{attribute 'external_name' := 'cmp_rts_DFC_rbr_safoutChnl3'}
TYPE DFC_rbr_safoutChnl3 : STRUCT
  DTC : UDINT := 16#200A00;
  DFCid : UINT := 802;
  debounceMethod : USINT := NO_DEBOUNCE;
END_STRUCT;
END_TYPE

{attribute 'external_name' := 'cmp_rts_DFC_rbr_safoutChnl4'}
TYPE DFC_rbr_safoutChnl4 : STRUCT
  DTC : UDINT := 16#200B00;
  DFCid : UINT := 805;
  debounceMethod : USINT := NO_DEBOUNCE;
END_STRUCT;
END_TYPE

{attribute 'external_name' := 'cmp_rts_DFC_rbr_safoutChnl5'}
TYPE DFC_rbr_safoutChnl5 : STRUCT
  DTC : UDINT := 16#200C00;
  DFCid : UINT := 808;
  debounceMethod : USINT := NO_DEBOUNCE;
END_STRUCT;
END_TYPE

{attribute 'external_name' := 'cmp_rts_DFC_rbr_safoutChnl6'}
TYPE DFC_rbr_safoutChnl6 : STRUCT
  DTC : UDINT := 16#201900;
  DFCid : UINT := 811;
  debounceMethod : USINT := NO_DEBOUNCE;
END_STRUCT;
END_TYPE

{attribute 'external_name' := 'cmp_rts_DFC_rbr_safoutChnl7'}
TYPE DFC_rbr_safoutChnl7 : STRUCT
  DTC : UDINT := 16#201A00;
  DFCid : UINT := 814;
  debounceMethod : USINT := NO_DEBOUNCE;
END_STRUCT;
END_TYPE

{attribute 'external_name' := 'cmp_rts_DFC_rbr_safoutChnl8'}
TYPE DFC_rbr_safoutChnl8 : STRUCT
  DTC : UDINT := 16#201B00;
  DFCid : UINT := 817;
  debounceMethod : USINT := NO_DEBOUNCE;
END_STRUCT;
END_TYPE

{attribute 'external_name' := 'cmp_rts_DFC_rbr_safoutChnl9'}
TYPE DFC_rbr_safoutChnl9 : STRUCT
  DTC : UDINT := 16#201C00;
  DFCid : UINT := 820;
  debounceMethod : USINT := NO_DEBOUNCE;
END_STRUCT;
END_TYPE

{attribute 'external_name' := 'cmp_rts_DFC_rbr_safoutChnl10'}
TYPE DFC_rbr_safoutChnl10 : STRUCT
  DTC : UDINT := 16#201D00;
  DFCid : UINT := 770;
  debounceMethod : USINT := NO_DEBOUNCE;
END_STRUCT;
END_TYPE

{attribute 'external_name' := 'cmp_rts_DFC_rbr_safoutChnl11'}
TYPE DFC_rbr_safoutChnl11 : STRUCT
  DTC : UDINT := 16#201E00;
  DFCid : UINT := 773;
  debounceMethod : USINT := NO_DEBOUNCE;
END_STRUCT;
END_TYPE

{attribute 'external_name' := 'cmp_rts_DFC_rbr_safoutChnl12'}
TYPE DFC_rbr_safoutChnl12 : STRUCT
  DTC : UDINT := 16#201F00;
  DFCid : UINT := 776;
  debounceMethod : USINT := NO_DEBOUNCE;
END_STRUCT;
END_TYPE

{attribute 'external_name' := 'cmp_rts_DFC_rbr_safoutChnl13'}
TYPE DFC_rbr_safoutChnl13 : STRUCT
  DTC : UDINT := 16#202000;
  DFCid : UINT := 779;
  debounceMethod : USINT := NO_DEBOUNCE;
END_STRUCT;
END_TYPE

{attribute 'external_name' := 'cmp_rts_DFC_rbr_safoutChnl14'}
TYPE DFC_rbr_safoutChnl14 : STRUCT
  DTC : UDINT := 16#202100;
  DFCid : UINT := 782;
  debounceMethod : USINT := NO_DEBOUNCE;
END_STRUCT;
END_TYPE

{attribute 'external_name' := 'cmp_rts_DFC_rbr_safoutChnl15'}
TYPE DFC_rbr_safoutChnl15 : STRUCT
  DTC : UDINT := 16#202200;
  DFCid : UINT := 785;
  debounceMethod : USINT := NO_DEBOUNCE;
END_STRUCT;
END_TYPE

{attribute 'external_name' := 'cmp_rts_DFC_rbr_safoutChnl16'}
TYPE DFC_rbr_safoutChnl16 : STRUCT
  DTC : UDINT := 16#202300;
  DFCid : UINT := 788;
  debounceMethod : USINT := NO_DEBOUNCE;
END_STRUCT;
END_TYPE

{attribute 'external_name' := 'cmp_rts_DFC_rbr_safoutChnl17'}
TYPE DFC_rbr_safoutChnl17 : STRUCT
  DTC : UDINT := 16#202400;
  DFCid : UINT := 791;
  debounceMethod : USINT := NO_DEBOUNCE;
END_STRUCT;
END_TYPE

{attribute 'external_name' := 'cmp_rts_DFC_rbr_safoutChnl18'}
TYPE DFC_rbr_safoutChnl18 : STRUCT
  DTC : UDINT := 16#202500;
  DFCid : UINT := 794;
  debounceMethod : USINT := NO_DEBOUNCE;
END_STRUCT;
END_TYPE

{attribute 'external_name' := 'cmp_rts_DFC_rbr_safoutChnl6Dev'}
TYPE DFC_rbr_safoutChnl6Dev : STRUCT
  DTC : UDINT := 16#202600;
  DFCid : UINT := 812;
  debounceMethod : USINT := NO_DEBOUNCE;
END_STRUCT;
END_TYPE

{attribute 'external_name' := 'cmp_rts_DFC_rbr_safoutChnl7Dev'}
TYPE DFC_rbr_safoutChnl7Dev : STRUCT
  DTC : UDINT := 16#202700;
  DFCid : UINT := 815;
  debounceMethod : USINT := NO_DEBOUNCE;
END_STRUCT;
END_TYPE

{attribute 'external_name' := 'cmp_rts_DFC_rbr_safoutChnl8Dev'}
TYPE DFC_rbr_safoutChnl8Dev : STRUCT
  DTC : UDINT := 16#202800;
  DFCid : UINT := 818;
  debounceMethod : USINT := NO_DEBOUNCE;
END_STRUCT;
END_TYPE

{attribute 'external_name' := 'cmp_rts_DFC_rbr_safoutChnl9Dev'}
TYPE DFC_rbr_safoutChnl9Dev : STRUCT
  DTC : UDINT := 16#202900;
  DFCid : UINT := 821;
  debounceMethod : USINT := NO_DEBOUNCE;
END_STRUCT;
END_TYPE

{attribute 'external_name' := 'cmp_rts_DFC_rbr_safoutChnl10Dev'}
TYPE DFC_rbr_safoutChnl10Dev : STRUCT
  DTC : UDINT := 16#202A00;
  DFCid : UINT := 771;
  debounceMethod : USINT := NO_DEBOUNCE;
END_STRUCT;
END_TYPE

{attribute 'external_name' := 'cmp_rts_DFC_rbr_safoutChnl11Dev'}
TYPE DFC_rbr_safoutChnl11Dev : STRUCT
  DTC : UDINT := 16#202B00;
  DFCid : UINT := 774;
  debounceMethod : USINT := NO_DEBOUNCE;
END_STRUCT;
END_TYPE

{attribute 'external_name' := 'cmp_rts_DFC_rbr_safoutChnl12Dev'}
TYPE DFC_rbr_safoutChnl12Dev : STRUCT
  DTC : UDINT := 16#202C00;
  DFCid : UINT := 777;
  debounceMethod : USINT := NO_DEBOUNCE;
END_STRUCT;
END_TYPE

{attribute 'external_name' := 'cmp_rts_DFC_rbr_safoutChnl13Dev'}
TYPE DFC_rbr_safoutChnl13Dev : STRUCT
  DTC : UDINT := 16#202D00;
  DFCid : UINT := 780;
  debounceMethod : USINT := NO_DEBOUNCE;
END_STRUCT;
END_TYPE

{attribute 'external_name' := 'cmp_rts_DFC_rbr_safoutChnl14Dev'}
TYPE DFC_rbr_safoutChnl14Dev : STRUCT
  DTC : UDINT := 16#202E00;
  DFCid : UINT := 783;
  debounceMethod : USINT := NO_DEBOUNCE;
END_STRUCT;
END_TYPE

{attribute 'external_name' := 'cmp_rts_DFC_rbr_safoutChnl15Dev'}
TYPE DFC_rbr_safoutChnl15Dev : STRUCT
  DTC : UDINT := 16#202F00;
  DFCid : UINT := 786;
  debounceMethod : USINT := NO_DEBOUNCE;
END_STRUCT;
END_TYPE

{attribute 'external_name' := 'cmp_rts_DFC_rbr_safoutChnl16Dev'}
TYPE DFC_rbr_safoutChnl16Dev : STRUCT
  DTC : UDINT := 16#203000;
  DFCid : UINT := 789;
  debounceMethod : USINT := NO_DEBOUNCE;
END_STRUCT;
END_TYPE

{attribute 'external_name' := 'cmp_rts_DFC_rbr_safoutChnl17Dev'}
TYPE DFC_rbr_safoutChnl17Dev : STRUCT
  DTC : UDINT := 16#203100;
  DFCid : UINT := 792;
  debounceMethod : USINT := NO_DEBOUNCE;
END_STRUCT;
END_TYPE

{attribute 'external_name' := 'cmp_rts_DFC_rbr_safoutChnl18Dev'}
TYPE DFC_rbr_safoutChnl18Dev : STRUCT
  DTC : UDINT := 16#203200;
  DFCid : UINT := 795;
  debounceMethod : USINT := NO_DEBOUNCE;
END_STRUCT;
END_TYPE

{attribute 'external_name' := 'cmp_rts_DFC_rbr_safoutChnl1OR'}
TYPE DFC_rbr_safoutChnl1OR : STRUCT
  DTC : UDINT := 16#200D00;
  DFCid : UINT := 798;
  debounceMethod : USINT := NO_DEBOUNCE;
END_STRUCT;
END_TYPE

{attribute 'external_name' := 'cmp_rts_DFC_rbr_safoutChnl2OR'}
TYPE DFC_rbr_safoutChnl2OR : STRUCT
  DTC : UDINT := 16#200E00;
  DFCid : UINT := 801;
  debounceMethod : USINT := NO_DEBOUNCE;
END_STRUCT;
END_TYPE

{attribute 'external_name' := 'cmp_rts_DFC_rbr_safoutChnl3OR'}
TYPE DFC_rbr_safoutChnl3OR : STRUCT
  DTC : UDINT := 16#200F00;
  DFCid : UINT := 804;
  debounceMethod : USINT := NO_DEBOUNCE;
END_STRUCT;
END_TYPE

{attribute 'external_name' := 'cmp_rts_DFC_rbr_safoutChnl4OR'}
TYPE DFC_rbr_safoutChnl4OR : STRUCT
  DTC : UDINT := 16#201100;
  DFCid : UINT := 807;
  debounceMethod : USINT := NO_DEBOUNCE;
END_STRUCT;
END_TYPE

{attribute 'external_name' := 'cmp_rts_DFC_rbr_safoutChnl5OR'}
TYPE DFC_rbr_safoutChnl5OR : STRUCT
  DTC : UDINT := 16#201200;
  DFCid : UINT := 810;
  debounceMethod : USINT := NO_DEBOUNCE;
END_STRUCT;
END_TYPE

{attribute 'external_name' := 'cmp_rts_DFC_rbr_safoutChnl6OR'}
TYPE DFC_rbr_safoutChnl6OR : STRUCT
  DTC : UDINT := 16#203300;
  DFCid : UINT := 813;
  debounceMethod : USINT := NO_DEBOUNCE;
END_STRUCT;
END_TYPE

{attribute 'external_name' := 'cmp_rts_DFC_rbr_safoutChnl7OR'}
TYPE DFC_rbr_safoutChnl7OR : STRUCT
  DTC : UDINT := 16#203400;
  DFCid : UINT := 816;
  debounceMethod : USINT := NO_DEBOUNCE;
END_STRUCT;
END_TYPE

{attribute 'external_name' := 'cmp_rts_DFC_rbr_safoutChnl8OR'}
TYPE DFC_rbr_safoutChnl8OR : STRUCT
  DTC : UDINT := 16#203500;
  DFCid : UINT := 819;
  debounceMethod : USINT := NO_DEBOUNCE;
END_STRUCT;
END_TYPE

{attribute 'external_name' := 'cmp_rts_DFC_rbr_safoutChnl9OR'}
TYPE DFC_rbr_safoutChnl9OR : STRUCT
  DTC : UDINT := 16#203600;
  DFCid : UINT := 822;
  debounceMethod : USINT := NO_DEBOUNCE;
END_STRUCT;
END_TYPE

{attribute 'external_name' := 'cmp_rts_DFC_rbr_safoutChnl10OR'}
TYPE DFC_rbr_safoutChnl10OR : STRUCT
  DTC : UDINT := 16#203700;
  DFCid : UINT := 772;
  debounceMethod : USINT := NO_DEBOUNCE;
END_STRUCT;
END_TYPE

{attribute 'external_name' := 'cmp_rts_DFC_rbr_safoutChnl11OR'}
TYPE DFC_rbr_safoutChnl11OR : STRUCT
  DTC : UDINT := 16#203800;
  DFCid : UINT := 775;
  debounceMethod : USINT := NO_DEBOUNCE;
END_STRUCT;
END_TYPE

{attribute 'external_name' := 'cmp_rts_DFC_rbr_safoutChnl12OR'}
TYPE DFC_rbr_safoutChnl12OR : STRUCT
  DTC : UDINT := 16#203900;
  DFCid : UINT := 778;
  debounceMethod : USINT := NO_DEBOUNCE;
END_STRUCT;
END_TYPE

{attribute 'external_name' := 'cmp_rts_DFC_rbr_safoutChnl13OR'}
TYPE DFC_rbr_safoutChnl13OR : STRUCT
  DTC : UDINT := 16#203A00;
  DFCid : UINT := 781;
  debounceMethod : USINT := NO_DEBOUNCE;
END_STRUCT;
END_TYPE

{attribute 'external_name' := 'cmp_rts_DFC_rbr_safoutChnl14OR'}
TYPE DFC_rbr_safoutChnl14OR : STRUCT
  DTC : UDINT := 16#203B00;
  DFCid : UINT := 784;
  debounceMethod : USINT := NO_DEBOUNCE;
END_STRUCT;
END_TYPE

{attribute 'external_name' := 'cmp_rts_DFC_rbr_safoutChnl15OR'}
TYPE DFC_rbr_safoutChnl15OR : STRUCT
  DTC : UDINT := 16#203C00;
  DFCid : UINT := 787;
  debounceMethod : USINT := NO_DEBOUNCE;
END_STRUCT;
END_TYPE

{attribute 'external_name' := 'cmp_rts_DFC_rbr_safoutChnl16OR'}
TYPE DFC_rbr_safoutChnl16OR : STRUCT
  DTC : UDINT := 16#203D00;
  DFCid : UINT := 790;
  debounceMethod : USINT := NO_DEBOUNCE;
END_STRUCT;
END_TYPE

{attribute 'external_name' := 'cmp_rts_DFC_rbr_safoutChnl17OR'}
TYPE DFC_rbr_safoutChnl17OR : STRUCT
  DTC : UDINT := 16#203E00;
  DFCid : UINT := 793;
  debounceMethod : USINT := NO_DEBOUNCE;
END_STRUCT;
END_TYPE

{attribute 'external_name' := 'cmp_rts_DFC_rbr_safoutChnl18OR'}
TYPE DFC_rbr_safoutChnl18OR : STRUCT
  DTC : UDINT := 16#203F00;
  DFCid : UINT := 796;
  debounceMethod : USINT := NO_DEBOUNCE;
END_STRUCT;
END_TYPE

{attribute 'external_name' := 'cmp_rts_DFC_rbr_safoutCfg'}
TYPE DFC_rbr_safoutCfg : STRUCT
  DTC : UDINT := 16#200100;
  DFCid : UINT := 768;
  debounceMethod : USINT := NO_DEBOUNCE;
END_STRUCT;
END_TYPE

{attribute 'external_name' := 'cmp_rts_DFC_rbr_safout'}
TYPE DFC_rbr_safout : STRUCT
  DTC : UDINT := 16#200200;
  DFCid : UINT := 767;
  debounceMethod : USINT := NO_DEBOUNCE;
END_STRUCT;
END_TYPE

{attribute 'external_name' := 'cmp_rts_DFC_rbr_safoutGetStatus'}
TYPE DFC_rbr_safoutGetStatus : STRUCT
  DTC : UDINT := 16#200300;
  DFCid : UINT := 824;
  debounceMethod : USINT := NO_DEBOUNCE;
END_STRUCT;
END_TYPE

{attribute 'external_name' := 'cmp_rts_DFC_rbr_safoutDevError'}
TYPE DFC_rbr_safoutDevError : STRUCT
  DTC : UDINT := 16#201800;
  DFCid : UINT := 823;
  debounceMethod : USINT := NO_DEBOUNCE;
END_STRUCT;
END_TYPE

{attribute 'external_name' := 'cmp_rts_DFC_rbr_safoutResetError'}
TYPE DFC_rbr_safoutResetError : STRUCT
  DTC : UDINT := 16#200400;
  DFCid : UINT := 826;
  debounceMethod : USINT := NO_DEBOUNCE;
END_STRUCT;
END_TYPE

{attribute 'external_name' := 'cmp_rts_DFC_rbr_safoutIgnoreError'}
TYPE DFC_rbr_safoutIgnoreError : STRUCT
  DTC : UDINT := 16#200500;
  DFCid : UINT := 825;
  debounceMethod : USINT := NO_DEBOUNCE;
END_STRUCT;
END_TYPE

{attribute 'external_name' := 'cmp_rts_DFC_rbr_safoutUnlock'}
TYPE DFC_rbr_safoutUnlock : STRUCT
  DTC : UDINT := 16#200600;
  DFCid : UINT := 827;
  debounceMethod : USINT := NO_DEBOUNCE;
END_STRUCT;
END_TYPE

{attribute 'external_name' := 'cmp_rts_DFC_rbr_outDo'}
TYPE DFC_rbr_outDo : STRUCT
  DTC : UDINT := 16#048300;
  DFCid : UINT := 721;
  debounceMethod : USINT := NO_DEBOUNCE;
END_STRUCT;
END_TYPE

{attribute 'external_name' := 'cmp_rts_DFC_rbr_outDoGetCurrent'}
TYPE DFC_rbr_outDoGetCurrent : STRUCT
  DTC : UDINT := 16#048400;
  DFCid : UINT := 724;
  debounceMethod : USINT := NO_DEBOUNCE;
END_STRUCT;
END_TYPE

{attribute 'external_name' := 'cmp_rts_DFC_rbr_outPod'}
TYPE DFC_rbr_outPod : STRUCT
  DTC : UDINT := 16#048B00;
  DFCid : UINT := 763;
  debounceMethod : USINT := NO_DEBOUNCE;
END_STRUCT;
END_TYPE

{attribute 'external_name' := 'cmp_rts_DFC_rbr_outPodCfg'}
TYPE DFC_rbr_outPodCfg : STRUCT
  DTC : UDINT := 16#048C00;
  DFCid : UINT := 764;
  debounceMethod : USINT := NO_DEBOUNCE;
END_STRUCT;
END_TYPE

{attribute 'external_name' := 'cmp_rts_DFC_rbr_outPodCfgPeriod'}
TYPE DFC_rbr_outPodCfgPeriod : STRUCT
  DTC : UDINT := 16#048D00;
  DFCid : UINT := 765;
  debounceMethod : USINT := NO_DEBOUNCE;
END_STRUCT;
END_TYPE

{attribute 'external_name' := 'cmp_rts_DFC_rbr_outPoc'}
TYPE DFC_rbr_outPoc : STRUCT
  DTC : UDINT := 16#048600;
  DFCid : UINT := 759;
  debounceMethod : USINT := NO_DEBOUNCE;
END_STRUCT;
END_TYPE

{attribute 'external_name' := 'cmp_rts_DFC_rbr_outPocCfg'}
TYPE DFC_rbr_outPocCfg : STRUCT
  DTC : UDINT := 16#048800;
  DFCid : UINT := 760;
  debounceMethod : USINT := NO_DEBOUNCE;
END_STRUCT;
END_TYPE

{attribute 'external_name' := 'cmp_rts_DFC_rbr_outPoCfg'}
TYPE DFC_rbr_outPoCfg : STRUCT
  DTC : UDINT := 16#048700;
  DFCid : UINT := 752;
  debounceMethod : USINT := NO_DEBOUNCE;
END_STRUCT;
END_TYPE

{attribute 'external_name' := 'cmp_rts_DFC_rbr_outPocCfgPI'}
TYPE DFC_rbr_outPocCfgPI : STRUCT
  DTC : UDINT := 16#048A00;
  DFCid : UINT := 762;
  debounceMethod : USINT := NO_DEBOUNCE;
END_STRUCT;
END_TYPE

{attribute 'external_name' := 'cmp_rts_DFC_rbr_outPocCfgDither'}
TYPE DFC_rbr_outPocCfgDither : STRUCT
  DTC : UDINT := 16#048900;
  DFCid : UINT := 761;
  debounceMethod : USINT := NO_DEBOUNCE;
END_STRUCT;
END_TYPE

{attribute 'external_name' := 'cmp_rts_DFC_rbr_outPoGetCurrent'}
TYPE DFC_rbr_outPoGetCurrent : STRUCT
  DTC : UDINT := 16#048E00;
  DFCid : UINT := 756;
  debounceMethod : USINT := NO_DEBOUNCE;
END_STRUCT;
END_TYPE

{attribute 'external_name' := 'cmp_rts_DFC_rbr_outAov'}
TYPE DFC_rbr_outAov : STRUCT
  DTC : UDINT := 16#048000;
  DFCid : UINT := 715;
  debounceMethod : USINT := NO_DEBOUNCE;
END_STRUCT;
END_TYPE

{attribute 'external_name' := 'cmp_rts_DFC_rbr_outAovCfg'}
TYPE DFC_rbr_outAovCfg : STRUCT
  DTC : UDINT := 16#048100;
  DFCid : UINT := 716;
  debounceMethod : USINT := NO_DEBOUNCE;
END_STRUCT;
END_TYPE

{attribute 'external_name' := 'cmp_rts_DFC_rbr_outAovCfgPI'}
TYPE DFC_rbr_outAovCfgPI : STRUCT
  DTC : UDINT := 16#14D700;
  DFCid : UINT := 717;
  debounceMethod : USINT := NO_DEBOUNCE;
END_STRUCT;
END_TYPE

{attribute 'external_name' := 'cmp_rts_DFC_rbr_outAovGetVoltage'}
TYPE DFC_rbr_outAovGetVoltage : STRUCT
  DTC : UDINT := 16#048200;
  DFCid : UINT := 719;
  debounceMethod : USINT := NO_DEBOUNCE;
END_STRUCT;
END_TYPE

{attribute 'external_name' := 'cmp_rts_DFC_rbr_outDoGetStatus'}
TYPE DFC_rbr_outDoGetStatus : STRUCT
  DTC : UDINT := 16#048F00;
  DFCid : UINT := 725;
  debounceMethod : USINT := NO_DEBOUNCE;
END_STRUCT;
END_TYPE

{attribute 'external_name' := 'cmp_rts_DFC_rbr_outDoResetError'}
TYPE DFC_rbr_outDoResetError : STRUCT
  DTC : UDINT := 16#049000;
  DFCid : UINT := 726;
  debounceMethod : USINT := NO_DEBOUNCE;
END_STRUCT;
END_TYPE

{attribute 'external_name' := 'cmp_rts_DFC_rbr_outPo'}
TYPE DFC_rbr_outPo : STRUCT
  DTC : UDINT := 16#049100;
  DFCid : UINT := 751;
  debounceMethod : USINT := NO_DEBOUNCE;
END_STRUCT;
END_TYPE

{attribute 'external_name' := 'cmp_rts_DFC_rbr_outPoCfgPeriod'}
TYPE DFC_rbr_outPoCfgPeriod : STRUCT
  DTC : UDINT := 16#049200;
  DFCid : UINT := 753;
  debounceMethod : USINT := NO_DEBOUNCE;
END_STRUCT;
END_TYPE

{attribute 'external_name' := 'cmp_rts_DFC_rbr_outPoGetStatus'}
TYPE DFC_rbr_outPoGetStatus : STRUCT
  DTC : UDINT := 16#049300;
  DFCid : UINT := 757;
  debounceMethod : USINT := NO_DEBOUNCE;
END_STRUCT;
END_TYPE

{attribute 'external_name' := 'cmp_rts_DFC_rbr_outPoResetError'}
TYPE DFC_rbr_outPoResetError : STRUCT
  DTC : UDINT := 16#049400;
  DFCid : UINT := 758;
  debounceMethod : USINT := NO_DEBOUNCE;
END_STRUCT;
END_TYPE

{attribute 'external_name' := 'cmp_rts_DFC_rbr_outAovGetStatus'}
TYPE DFC_rbr_outAovGetStatus : STRUCT
  DTC : UDINT := 16#049500;
  DFCid : UINT := 718;
  debounceMethod : USINT := NO_DEBOUNCE;
END_STRUCT;
END_TYPE

{attribute 'external_name' := 'cmp_rts_DFC_rbr_outAovResetError'}
TYPE DFC_rbr_outAovResetError : STRUCT
  DTC : UDINT := 16#049600;
  DFCid : UINT := 720;
  debounceMethod : USINT := NO_DEBOUNCE;
END_STRUCT;
END_TYPE

{attribute 'external_name' := 'cmp_rts_DFC_rbr_sysAiv'}
TYPE DFC_rbr_sysAiv : STRUCT
  DTC : UDINT := 16#010100;
  DFCid : UINT := 842;
  debounceMethod : USINT := NO_DEBOUNCE;
END_STRUCT;
END_TYPE

{attribute 'external_name' := 'cmp_rts_DFC_rbr_memFlsCfgShr'}
TYPE DFC_rbr_memFlsCfgShr : STRUCT
  DTC : UDINT := 16#060900;
  DFCid : UINT := 649;
  debounceMethod : USINT := NO_DEBOUNCE;
END_STRUCT;
END_TYPE

{attribute 'external_name' := 'cmp_rts_DFC_rbr_sysDo'}
TYPE DFC_rbr_sysDo : STRUCT
  DTC : UDINT := 16#010200;
  DFCid : UINT := 844;
  debounceMethod : USINT := NO_DEBOUNCE;
END_STRUCT;
END_TYPE

{attribute 'external_name' := 'cmp_rts_DFC_rbr_sysGetVss'}
TYPE DFC_rbr_sysGetVss : STRUCT
  DTC : UDINT := 16#010600;
  DFCid : UINT := 845;
  debounceMethod : USINT := NO_DEBOUNCE;
END_STRUCT;
END_TYPE

{attribute 'external_name' := 'cmp_rts_DFC_rbr_sysDi'}
TYPE DFC_rbr_sysDi : STRUCT
  DTC : UDINT := 16#010300;
  DFCid : UINT := 843;
  debounceMethod : USINT := NO_DEBOUNCE;
END_STRUCT;
END_TYPE

{attribute 'external_name' := 'cmp_rts_DFC_rbr_sysAit'}
TYPE DFC_rbr_sysAit : STRUCT
  DTC : UDINT := 16#010400;
  DFCid : UINT := 841;
  debounceMethod : USINT := NO_DEBOUNCE;
END_STRUCT;
END_TYPE

{attribute 'external_name' := 'cmp_rts_DFC_rbr_sysSetVss'}
TYPE DFC_rbr_sysSetVss : STRUCT
  DTC : UDINT := 16#010500;
  DFCid : UINT := 849;
  debounceMethod : USINT := NO_DEBOUNCE;
END_STRUCT;
END_TYPE

{attribute 'external_name' := 'cmp_rts_DFC_rbr_outPoDisable'}
TYPE DFC_rbr_outPoDisable : STRUCT
  DTC : UDINT := 16#049800;
  DFCid : UINT := 755;
  debounceMethod : USINT := NO_DEBOUNCE;
END_STRUCT;
END_TYPE

{attribute 'external_name' := 'cmp_rts_DFC_rbr_safout_cfgDiag'}
TYPE DFC_rbr_safout_cfgDiag : STRUCT
  DTC : UDINT := 16#200700;
  DFCid : UINT := 828;
  debounceMethod : USINT := NO_DEBOUNCE;
END_STRUCT;
END_TYPE

{attribute 'external_name' := 'cmp_rts_DFC_rbr_outDoDisable'}
TYPE DFC_rbr_outDoDisable : STRUCT
  DTC : UDINT := 16#049700;
  DFCid : UINT := 723;
  debounceMethod : USINT := NO_DEBOUNCE;
END_STRUCT;
END_TYPE

{attribute 'external_name' := 'cmp_rts_DFC_rbr_sysOperHrIntegrityErr'}
TYPE DFC_rbr_sysOperHrIntegrityErr : STRUCT
  DTC : UDINT := 16#010A00;
  DFCid : UINT := 847;
  debounceMethod : USINT := NO_DEBOUNCE;
END_STRUCT;
END_TYPE

{attribute 'external_name' := 'cmp_rts_DFC_rbr_sysOperHrsSaturated'}
TYPE DFC_rbr_sysOperHrsSaturated : STRUCT
  DTC : UDINT := 16#010B00;
  DFCid : UINT := 848;
  debounceMethod : USINT := NO_DEBOUNCE;
END_STRUCT;
END_TYPE

{attribute 'external_name' := 'cmp_rts_DFC_rbr_mo_INHLatch'}
TYPE DFC_rbr_mo_INHLatch : STRUCT
  DTC : UDINT := 16#082200;
  DFCid : UINT := 664;
  debounceMethod : USINT := NO_DEBOUNCE;
END_STRUCT;
END_TYPE

{attribute 'external_name' := 'cmp_rts_DFC_rbr_rsmFfiApiCallErr'}
TYPE DFC_rbr_rsmFfiApiCallErr : STRUCT
  DTC : UDINT := 16#010C00;
  DFCid : UINT := 766;
  debounceMethod : USINT := NO_DEBOUNCE;
END_STRUCT;
END_TYPE

{attribute 'external_name' := 'cmp_rts_DFC_rbr_mo_INH'}
TYPE DFC_rbr_mo_INH : STRUCT
  DTC : UDINT := 16#082100;
  DFCid : UINT := 663;
  debounceMethod : USINT := NO_DEBOUNCE;
END_STRUCT;
END_TYPE

{attribute 'external_name' := 'cmp_rts_DFC_rbr_memReadSystemError'}
TYPE DFC_rbr_memReadSystemError : STRUCT
  DTC : UDINT := 16#060800;
  DFCid : UINT := 657;
  debounceMethod : USINT := NO_DEBOUNCE;
END_STRUCT;
END_TYPE

{attribute 'external_name' := 'cmp_rts_DFC_rbr_memReadCalibInputError'}
TYPE DFC_rbr_memReadCalibInputError : STRUCT
  DTC : UDINT := 16#060A00;
  DFCid : UINT := 655;
  debounceMethod : USINT := NO_DEBOUNCE;
END_STRUCT;
END_TYPE

{attribute 'external_name' := 'cmp_rts_DFC_rbr_memReadCalibOuputError'}
TYPE DFC_rbr_memReadCalibOuputError : STRUCT
  DTC : UDINT := 16#060B00;
  DFCid : UINT := 656;
  debounceMethod : USINT := NO_DEBOUNCE;
END_STRUCT;
END_TYPE

{attribute 'external_name' := 'cmp_rts_DFC_rbr_memReadApi2Error'}
TYPE DFC_rbr_memReadApi2Error : STRUCT
  DTC : UDINT := 16#060600;
  DFCid : UINT := 653;
  debounceMethod : USINT := NO_DEBOUNCE;
END_STRUCT;
END_TYPE

{attribute 'external_name' := 'cmp_rts_DFC_rbr_memReadApi1Error'}
TYPE DFC_rbr_memReadApi1Error : STRUCT
  DTC : UDINT := 16#060500;
  DFCid : UINT := 652;
  debounceMethod : USINT := NO_DEBOUNCE;
END_STRUCT;
END_TYPE

{attribute 'external_name' := 'cmp_rts_DFC_rbr_memMarkBlock'}
TYPE DFC_rbr_memMarkBlock : STRUCT
  DTC : UDINT := 16#060400;
  DFCid : UINT := 651;
  debounceMethod : USINT := NO_DEBOUNCE;
END_STRUCT;
END_TYPE

{attribute 'external_name' := 'cmp_rts_DFC_rbr_safoutChnl3Dev'}
TYPE DFC_rbr_safoutChnl3Dev : STRUCT
  DTC : UDINT := 16#201500;
  DFCid : UINT := 803;
  debounceMethod : USINT := NO_DEBOUNCE;
END_STRUCT;
END_TYPE

{attribute 'external_name' := 'cmp_rts_DFC_rbr_safoutChnl5Dev'}
TYPE DFC_rbr_safoutChnl5Dev : STRUCT
  DTC : UDINT := 16#201700;
  DFCid : UINT := 809;
  debounceMethod : USINT := NO_DEBOUNCE;
END_STRUCT;
END_TYPE

{attribute 'external_name' := 'cmp_rts_DFC_rbr_safoutChnl4Dev'}
TYPE DFC_rbr_safoutChnl4Dev : STRUCT
  DTC : UDINT := 16#201600;
  DFCid : UINT := 806;
  debounceMethod : USINT := NO_DEBOUNCE;
END_STRUCT;
END_TYPE

{attribute 'external_name' := 'cmp_rts_DFC_rbr_safoutChnl2Dev'}
TYPE DFC_rbr_safoutChnl2Dev : STRUCT
  DTC : UDINT := 16#201400;
  DFCid : UINT := 800;
  debounceMethod : USINT := NO_DEBOUNCE;
END_STRUCT;
END_TYPE

{attribute 'external_name' := 'cmp_rts_DFC_rbr_safoutChnl1Dev'}
TYPE DFC_rbr_safoutChnl1Dev : STRUCT
  DTC : UDINT := 16#201300;
  DFCid : UINT := 797;
  debounceMethod : USINT := NO_DEBOUNCE;
END_STRUCT;
END_TYPE

{attribute 'external_name' := 'cmp_rts_DFC_rbr_outDoCfgPwrLs'}
TYPE DFC_rbr_outDoCfgPwrLs : STRUCT
  DTC : UDINT := 16#14D800;
  DFCid : UINT := 722;
  debounceMethod : USINT := NO_DEBOUNCE;
END_STRUCT;
END_TYPE

{attribute 'external_name' := 'cmp_rts_DFC_rbr_outPoCfgPwrLs'}
TYPE DFC_rbr_outPoCfgPwrLs : STRUCT
  DTC : UDINT := 16#049900;
  DFCid : UINT := 754;
  debounceMethod : USINT := NO_DEBOUNCE;
END_STRUCT;
END_TYPE

{attribute 'external_name' := 'cmp_rts_DFC_rbr_lin_wakeUp'}
TYPE DFC_rbr_lin_wakeUp : STRUCT
  DTC : UDINT := 16#210000;
  DFCid : UINT := 648;
  debounceMethod : USINT := NO_DEBOUNCE;
END_STRUCT;
END_TYPE

{attribute 'external_name' := 'cmp_rts_DFC_rbr_lin_gotoSleep'}
TYPE DFC_rbr_lin_gotoSleep : STRUCT
  DTC : UDINT := 16#210200;
  DFCid : UINT := 646;
  debounceMethod : USINT := NO_DEBOUNCE;
END_STRUCT;
END_TYPE

{attribute 'external_name' := 'cmp_rts_DFC_rbr_lin_getStatus'}
TYPE DFC_rbr_lin_getStatus : STRUCT
  DTC : UDINT := 16#210300;
  DFCid : UINT := 645;
  debounceMethod : USINT := NO_DEBOUNCE;
END_STRUCT;
END_TYPE

{attribute 'external_name' := 'cmp_rts_DFC_rbr_lin_scheduleRequest'}
TYPE DFC_rbr_lin_scheduleRequest : STRUCT
  DTC : UDINT := 16#210100;
  DFCid : UINT := 647;
  debounceMethod : USINT := NO_DEBOUNCE;
END_STRUCT;
END_TYPE

{attribute 'external_name' := 'cmp_rts_DFC_rbr_lin_SendSignal'}
TYPE DFC_rbr_lin_SendSignal : STRUCT
  DTC : UDINT := 16#210400;
  DFCid : UINT := 644;
  debounceMethod : USINT := NO_DEBOUNCE;
END_STRUCT;
END_TYPE

{attribute 'external_name' := 'cmp_rts_DFC_rbr_inPhaseGetStatus'}
TYPE DFC_rbr_inPhaseGetStatus : STRUCT
  DTC : UDINT := 16#039F00;
  DFCid : UINT := 593;
  debounceMethod : USINT := NO_DEBOUNCE;
END_STRUCT;
END_TYPE

{attribute 'external_name' := 'cmp_rts_DFC_rbr_inPhaseResetCounter'}
TYPE DFC_rbr_inPhaseResetCounter : STRUCT
  DTC : UDINT := 16#03A000;
  DFCid : UINT := 594;
  debounceMethod : USINT := NO_DEBOUNCE;
END_STRUCT;
END_TYPE

{attribute 'external_name' := 'cmp_rts_DFC_rbr_inPhase'}
TYPE DFC_rbr_inPhase : STRUCT
  DTC : UDINT := 16#039E00;
  DFCid : UINT := 592;
  debounceMethod : USINT := NO_DEBOUNCE;
END_STRUCT;
END_TYPE

{attribute 'external_name' := 'cmp_rts_DFC_rbr_inFi_Buffered'}
TYPE DFC_rbr_inFi_Buffered : STRUCT
  DTC : UDINT := 16#135200;
  DFCid : UINT := 591;
  debounceMethod : USINT := NO_DEBOUNCE;
END_STRUCT;
END_TYPE

{attribute 'external_name' := 'cmp_rts_DFC_rbr_secGetLevel'}
TYPE DFC_rbr_secGetLevel : STRUCT
  DTC : UDINT := 16#220200;
  DFCid : UINT := 833;
  debounceMethod : USINT := NO_DEBOUNCE;
END_STRUCT;
END_TYPE

{attribute 'external_name' := 'cmp_rts_DFC_rbr_secSetLevel'}
TYPE DFC_rbr_secSetLevel : STRUCT
  DTC : UDINT := 16#220300;
  DFCid : UINT := 840;
  debounceMethod : USINT := NO_DEBOUNCE;
END_STRUCT;
END_TYPE

{attribute 'external_name' := 'cmp_rts_DFC_rbr_secSaveSecret'}
TYPE DFC_rbr_secSaveSecret : STRUCT
  DTC : UDINT := 16#220100;
  DFCid : UINT := 839;
  debounceMethod : USINT := NO_DEBOUNCE;
END_STRUCT;
END_TYPE

{attribute 'external_name' := 'cmp_rts_DFC_rbr_secGetSeed'}
TYPE DFC_rbr_secGetSeed : STRUCT
  DTC : UDINT := 16#220000;
  DFCid : UINT := 835;
  debounceMethod : USINT := NO_DEBOUNCE;
END_STRUCT;
END_TYPE

{attribute 'external_name' := 'cmp_rts_DFC_rbr_secIsRequestAllowed'}
TYPE DFC_rbr_secIsRequestAllowed : STRUCT
  DTC : UDINT := 16#220700;
  DFCid : UINT := 837;
  debounceMethod : USINT := NO_DEBOUNCE;
END_STRUCT;
END_TYPE

{attribute 'external_name' := 'cmp_rts_DFC_rbr_secGetRnd'}
TYPE DFC_rbr_secGetRnd : STRUCT
  DTC : UDINT := 16#220600;
  DFCid : UINT := 834;
  debounceMethod : USINT := NO_DEBOUNCE;
END_STRUCT;
END_TYPE

{attribute 'external_name' := 'cmp_rts_DFC_rbr_secEvalRespKey'}
TYPE DFC_rbr_secEvalRespKey : STRUCT
  DTC : UDINT := 16#220500;
  DFCid : UINT := 831;
  debounceMethod : USINT := NO_DEBOUNCE;
END_STRUCT;
END_TYPE

{attribute 'external_name' := 'cmp_rts_DFC_rbr_secAccessDenied_RC'}
TYPE DFC_rbr_secAccessDenied_RC : STRUCT
  DTC : UDINT := 16#220B00;
  DFCid : UINT := 829;
  debounceMethod : USINT := NO_DEBOUNCE;
END_STRUCT;
END_TYPE

{attribute 'external_name' := 'cmp_rts_DFC_rbr_secAccessDenied_WDBI'}
TYPE DFC_rbr_secAccessDenied_WDBI : STRUCT
  DTC : UDINT := 16#220A00;
  DFCid : UINT := 830;
  debounceMethod : USINT := NO_DEBOUNCE;
END_STRUCT;
END_TYPE

{attribute 'external_name' := 'cmp_rts_DFC_rbr_secFlashingFailure'}
TYPE DFC_rbr_secFlashingFailure : STRUCT
  DTC : UDINT := 16#220900;
  DFCid : UINT := 832;
  debounceMethod : USINT := NO_DEBOUNCE;
END_STRUCT;
END_TYPE

{attribute 'external_name' := 'cmp_rts_DFC_rbr_secInvalidPassword'}
TYPE DFC_rbr_secInvalidPassword : STRUCT
  DTC : UDINT := 16#220800;
  DFCid : UINT := 836;
  debounceMethod : USINT := NO_DEBOUNCE;
END_STRUCT;
END_TYPE

{attribute 'external_name' := 'cmp_rts_DFC_rbr_secResetLevel'}
TYPE DFC_rbr_secResetLevel : STRUCT
  DTC : UDINT := 16#220400;
  DFCid : UINT := 838;
  debounceMethod : USINT := NO_DEBOUNCE;
END_STRUCT;
END_TYPE

{attribute 'external_name' := 'cmp_rts_DFC_rbr_lin_ReceiveSignal'}
TYPE DFC_rbr_lin_ReceiveSignal : STRUCT
  DTC : UDINT := 16#210500;
  DFCid : UINT := 643;
  debounceMethod : USINT := NO_DEBOUNCE;
END_STRUCT;
END_TYPE

{attribute 'external_name' := 'cmp_rts_DFC_rbr_sys_coreload'}
TYPE DFC_rbr_sys_coreload : STRUCT
  DTC : UDINT := 16#010900;
  DFCid : UINT := 850;
  debounceMethod : USINT := NO_DEBOUNCE;
END_STRUCT;
END_TYPE

{attribute 'external_name' := 'cmp_rts_DFC_rbr_sys_taskload'}
TYPE DFC_rbr_sys_taskload : STRUCT
  DTC : UDINT := 16#010800;
  DFCid : UINT := 851;
  debounceMethod : USINT := NO_DEBOUNCE;
END_STRUCT;
END_TYPE

{attribute 'external_name' := 'cmp_rts_DFC_rbr_dsmDTCJ1939'}
TYPE DFC_rbr_dsmDTCJ1939 : STRUCT
  DTC : UDINT := 16#071000;
  DFCid : UINT := 564;
  debounceMethod : USINT := NO_DEBOUNCE;
END_STRUCT;
END_TYPE

{attribute 'external_name' := 'cmp_rts_DFC_rbr_sysInit'}
TYPE DFC_rbr_sysInit : STRUCT
  DTC : UDINT := 16#010700;
  DFCid : UINT := 846;
  debounceMethod : USINT := NO_DEBOUNCE;
END_STRUCT;
END_TYPE

{attribute 'external_name' := 'cmp_rts_DFC_rbr_outK07Unintended'}
TYPE DFC_rbr_outK07Unintended : STRUCT
  DTC : UDINT := 16#14CB00;
  DFCid : UINT := 728;
  debounceMethod : USINT := NO_DEBOUNCE;
END_STRUCT;
END_TYPE

{attribute 'external_name' := 'cmp_rts_DFC_rbr_outK09Unintended'}
TYPE DFC_rbr_outK09Unintended : STRUCT
  DTC : UDINT := 16#14CD00;
  DFCid : UINT := 732;
  debounceMethod : USINT := NO_DEBOUNCE;
END_STRUCT;
END_TYPE

{attribute 'external_name' := 'cmp_rts_DFC_rbr_outK73Unintended'}
TYPE DFC_rbr_outK73Unintended : STRUCT
  DTC : UDINT := 16#14D600;
  DFCid : UINT := 750;
  debounceMethod : USINT := NO_DEBOUNCE;
END_STRUCT;
END_TYPE

{attribute 'external_name' := 'cmp_rts_DFC_rbr_outK08Unintended'}
TYPE DFC_rbr_outK08Unintended : STRUCT
  DTC : UDINT := 16#14CC00;
  DFCid : UINT := 730;
  debounceMethod : USINT := NO_DEBOUNCE;
END_STRUCT;
END_TYPE

{attribute 'external_name' := 'cmp_rts_DFC_rbr_outK29Unintended'}
TYPE DFC_rbr_outK29Unintended : STRUCT
  DTC : UDINT := 16#14D400;
  DFCid : UINT := 746;
  debounceMethod : USINT := NO_DEBOUNCE;
END_STRUCT;
END_TYPE

{attribute 'external_name' := 'cmp_rts_DFC_rbr_outK17Unintended'}
TYPE DFC_rbr_outK17Unintended : STRUCT
  DTC : UDINT := 16#14D300;
  DFCid : UINT := 744;
  debounceMethod : USINT := NO_DEBOUNCE;
END_STRUCT;
END_TYPE

{attribute 'external_name' := 'cmp_rts_DFC_rbr_outK16Unintended'}
TYPE DFC_rbr_outK16Unintended : STRUCT
  DTC : UDINT := 16#14D200;
  DFCid : UINT := 742;
  debounceMethod : USINT := NO_DEBOUNCE;
END_STRUCT;
END_TYPE

{attribute 'external_name' := 'cmp_rts_DFC_rbr_outK14Unintended'}
TYPE DFC_rbr_outK14Unintended : STRUCT
  DTC : UDINT := 16#14D000;
  DFCid : UINT := 738;
  debounceMethod : USINT := NO_DEBOUNCE;
END_STRUCT;
END_TYPE

{attribute 'external_name' := 'cmp_rts_DFC_rbr_outK15Unintended'}
TYPE DFC_rbr_outK15Unintended : STRUCT
  DTC : UDINT := 16#14D100;
  DFCid : UINT := 740;
  debounceMethod : USINT := NO_DEBOUNCE;
END_STRUCT;
END_TYPE

{attribute 'external_name' := 'cmp_rts_DFC_rbr_outK51Unintended'}
TYPE DFC_rbr_outK51Unintended : STRUCT
  DTC : UDINT := 16#14D500;
  DFCid : UINT := 748;
  debounceMethod : USINT := NO_DEBOUNCE;
END_STRUCT;
END_TYPE

{attribute 'external_name' := 'cmp_rts_DFC_rbr_outK12Unintended'}
TYPE DFC_rbr_outK12Unintended : STRUCT
  DTC : UDINT := 16#14CE00;
  DFCid : UINT := 734;
  debounceMethod : USINT := NO_DEBOUNCE;
END_STRUCT;
END_TYPE

{attribute 'external_name' := 'cmp_rts_DFC_rbr_outK13Unintended'}
TYPE DFC_rbr_outK13Unintended : STRUCT
  DTC : UDINT := 16#14CF00;
  DFCid : UINT := 736;
  debounceMethod : USINT := NO_DEBOUNCE;
END_STRUCT;
END_TYPE

{attribute 'external_name' := 'cmp_rts_DFC_rbr_outA32Unintended'}
TYPE DFC_rbr_outA32Unintended : STRUCT
  DTC : UDINT := 16#14C000;
  DFCid : UINT := 694;
  debounceMethod : USINT := NO_DEBOUNCE;
END_STRUCT;
END_TYPE

{attribute 'external_name' := 'cmp_rts_DFC_rbr_outA47Unintended'}
TYPE DFC_rbr_outA47Unintended : STRUCT
  DTC : UDINT := 16#14C500;
  DFCid : UINT := 704;
  debounceMethod : USINT := NO_DEBOUNCE;
END_STRUCT;
END_TYPE

{attribute 'external_name' := 'cmp_rts_DFC_rbr_outA31Unintended'}
TYPE DFC_rbr_outA31Unintended : STRUCT
  DTC : UDINT := 16#14BF00;
  DFCid : UINT := 692;
  debounceMethod : USINT := NO_DEBOUNCE;
END_STRUCT;
END_TYPE

{attribute 'external_name' := 'cmp_rts_DFC_rbr_outA48Unintended'}
TYPE DFC_rbr_outA48Unintended : STRUCT
  DTC : UDINT := 16#14C600;
  DFCid : UINT := 706;
  debounceMethod : USINT := NO_DEBOUNCE;
END_STRUCT;
END_TYPE

{attribute 'external_name' := 'cmp_rts_DFC_rbr_outA46Unintended'}
TYPE DFC_rbr_outA46Unintended : STRUCT
  DTC : UDINT := 16#14C400;
  DFCid : UINT := 702;
  debounceMethod : USINT := NO_DEBOUNCE;
END_STRUCT;
END_TYPE

{attribute 'external_name' := 'cmp_rts_DFC_rbr_outA33Unintended'}
TYPE DFC_rbr_outA33Unintended : STRUCT
  DTC : UDINT := 16#14C100;
  DFCid : UINT := 696;
  debounceMethod : USINT := NO_DEBOUNCE;
END_STRUCT;
END_TYPE

{attribute 'external_name' := 'cmp_rts_DFC_rbr_outA19Unintended'}
TYPE DFC_rbr_outA19Unintended : STRUCT
  DTC : UDINT := 16#14BD00;
  DFCid : UINT := 688;
  debounceMethod : USINT := NO_DEBOUNCE;
END_STRUCT;
END_TYPE

{attribute 'external_name' := 'cmp_rts_DFC_rbr_outA05Unintended'}
TYPE DFC_rbr_outA05Unintended : STRUCT
  DTC : UDINT := 16#14B600;
  DFCid : UINT := 674;
  debounceMethod : USINT := NO_DEBOUNCE;
END_STRUCT;
END_TYPE

{attribute 'external_name' := 'cmp_rts_DFC_rbr_outA20Unintended'}
TYPE DFC_rbr_outA20Unintended : STRUCT
  DTC : UDINT := 16#14BE00;
  DFCid : UINT := 690;
  debounceMethod : USINT := NO_DEBOUNCE;
END_STRUCT;
END_TYPE

{attribute 'external_name' := 'cmp_rts_DFC_rbr_outA03Unintended'}
TYPE DFC_rbr_outA03Unintended : STRUCT
  DTC : UDINT := 16#14B400;
  DFCid : UINT := 670;
  debounceMethod : USINT := NO_DEBOUNCE;
END_STRUCT;
END_TYPE

{attribute 'external_name' := 'cmp_rts_DFC_rbr_outA18Unintended'}
TYPE DFC_rbr_outA18Unintended : STRUCT
  DTC : UDINT := 16#14BC00;
  DFCid : UINT := 686;
  debounceMethod : USINT := NO_DEBOUNCE;
END_STRUCT;
END_TYPE

{attribute 'external_name' := 'cmp_rts_DFC_rbr_outA04Unintended'}
TYPE DFC_rbr_outA04Unintended : STRUCT
  DTC : UDINT := 16#14B500;
  DFCid : UINT := 672;
  debounceMethod : USINT := NO_DEBOUNCE;
END_STRUCT;
END_TYPE

{attribute 'external_name' := 'cmp_rts_DFC_rbr_outA34Unintended'}
TYPE DFC_rbr_outA34Unintended : STRUCT
  DTC : UDINT := 16#14C200;
  DFCid : UINT := 698;
  debounceMethod : USINT := NO_DEBOUNCE;
END_STRUCT;
END_TYPE

{attribute 'external_name' := 'cmp_rts_DFC_rbr_outA51Unintended'}
TYPE DFC_rbr_outA51Unintended : STRUCT
  DTC : UDINT := 16#14C700;
  DFCid : UINT := 708;
  debounceMethod : USINT := NO_DEBOUNCE;
END_STRUCT;
END_TYPE

{attribute 'external_name' := 'cmp_rts_DFC_rbr_outA35Unintended'}
TYPE DFC_rbr_outA35Unintended : STRUCT
  DTC : UDINT := 16#14C300;
  DFCid : UINT := 700;
  debounceMethod : USINT := NO_DEBOUNCE;
END_STRUCT;
END_TYPE

{attribute 'external_name' := 'cmp_rts_DFC_rbr_outA53Unintended'}
TYPE DFC_rbr_outA53Unintended : STRUCT
  DTC : UDINT := 16#14C900;
  DFCid : UINT := 712;
  debounceMethod : USINT := NO_DEBOUNCE;
END_STRUCT;
END_TYPE

{attribute 'external_name' := 'cmp_rts_DFC_rbr_outA52Unintended'}
TYPE DFC_rbr_outA52Unintended : STRUCT
  DTC : UDINT := 16#14C800;
  DFCid : UINT := 710;
  debounceMethod : USINT := NO_DEBOUNCE;
END_STRUCT;
END_TYPE

{attribute 'external_name' := 'cmp_rts_DFC_rbr_outA54Unintended'}
TYPE DFC_rbr_outA54Unintended : STRUCT
  DTC : UDINT := 16#14CA00;
  DFCid : UINT := 714;
  debounceMethod : USINT := NO_DEBOUNCE;
END_STRUCT;
END_TYPE

{attribute 'external_name' := 'cmp_rts_DFC_rbr_outA09Unintended'}
TYPE DFC_rbr_outA09Unintended : STRUCT
  DTC : UDINT := 16#14B900;
  DFCid : UINT := 680;
  debounceMethod : USINT := NO_DEBOUNCE;
END_STRUCT;
END_TYPE

{attribute 'external_name' := 'cmp_rts_DFC_rbr_outA02Unintended'}
TYPE DFC_rbr_outA02Unintended : STRUCT
  DTC : UDINT := 16#14B300;
  DFCid : UINT := 668;
  debounceMethod : USINT := NO_DEBOUNCE;
END_STRUCT;
END_TYPE

{attribute 'external_name' := 'cmp_rts_DFC_rbr_outA17Unintended'}
TYPE DFC_rbr_outA17Unintended : STRUCT
  DTC : UDINT := 16#14BB00;
  DFCid : UINT := 684;
  debounceMethod : USINT := NO_DEBOUNCE;
END_STRUCT;
END_TYPE

{attribute 'external_name' := 'cmp_rts_DFC_rbr_outA08Unintended'}
TYPE DFC_rbr_outA08Unintended : STRUCT
  DTC : UDINT := 16#14B800;
  DFCid : UINT := 678;
  debounceMethod : USINT := NO_DEBOUNCE;
END_STRUCT;
END_TYPE

{attribute 'external_name' := 'cmp_rts_DFC_rbr_outA07Unintended'}
TYPE DFC_rbr_outA07Unintended : STRUCT
  DTC : UDINT := 16#14B700;
  DFCid : UINT := 676;
  debounceMethod : USINT := NO_DEBOUNCE;
END_STRUCT;
END_TYPE

{attribute 'external_name' := 'cmp_rts_DFC_rbr_outA10Unintended'}
TYPE DFC_rbr_outA10Unintended : STRUCT
  DTC : UDINT := 16#14BA00;
  DFCid : UINT := 682;
  debounceMethod : USINT := NO_DEBOUNCE;
END_STRUCT;
END_TYPE

{attribute 'external_name' := 'cmp_rts_DFC_rbr_isobusSftyCanTxErr'}
TYPE DFC_rbr_isobusSftyCanTxErr : STRUCT
  DTC : UDINT := 16#051F00;
  DFCid : UINT := 642;
  debounceMethod : USINT := NO_DEBOUNCE;
END_STRUCT;
END_TYPE

{attribute 'external_name' := 'cmp_rts_DFC_rbr_dsmInitQueueOverflow'}
TYPE DFC_rbr_dsmInitQueueOverflow : STRUCT
  DTC : UDINT := 16#071400;
  DFCid : UINT := 571;
  debounceMethod : USINT := NO_DEBOUNCE;
END_STRUCT;
END_TYPE

{attribute 'external_name' := 'cmp_rts_DFC_rbr_mo_UV_VSS2'}
TYPE DFC_rbr_mo_UV_VSS2 : STRUCT
  DTC : UDINT := 16#080400;
  DFCid : UINT := 855;
  debounceMethod : USINT := NO_DEBOUNCE;
END_STRUCT;
END_TYPE

{attribute 'external_name' := 'cmp_rts_DFC_rbr_mo_UV_VSS1'}
TYPE DFC_rbr_mo_UV_VSS1 : STRUCT
  DTC : UDINT := 16#080200;
  DFCid : UINT := 854;
  debounceMethod : USINT := NO_DEBOUNCE;
END_STRUCT;
END_TYPE

{attribute 'external_name' := 'cmp_rts_DFC_rbr_mo_OV_VSS2'}
TYPE DFC_rbr_mo_OV_VSS2 : STRUCT
  DTC : UDINT := 16#080300;
  DFCid : UINT := 853;
  debounceMethod : USINT := NO_DEBOUNCE;
END_STRUCT;
END_TYPE

{attribute 'external_name' := 'cmp_rts_DFC_rbr_mo_OV_VSS1'}
TYPE DFC_rbr_mo_OV_VSS1 : STRUCT
  DTC : UDINT := 16#080100;
  DFCid : UINT := 852;
  debounceMethod : USINT := NO_DEBOUNCE;
END_STRUCT;
END_TYPE

{attribute 'external_name' := 'cmp_rts_DFC_ComCntESP_05'}
TYPE DFC_ComCntESP_05 : STRUCT
  DTC : UDINT := 16#102200;
END_STRUCT;
END_TYPE

{attribute 'external_name' := 'cmp_rts_DFC_MOXEMM_SMU_ALM3_1'}
TYPE DFC_MOXEMM_SMU_ALM3_1 : STRUCT
  DTC : UDINT := 16#108800;
  DFCid : UINT := 933;
  debounceMethod : USINT := NATIVE;
END_STRUCT;
END_TYPE

{attribute 'external_name' := 'cmp_rts_DFC_MOXEMM_SMU_ALM3_2'}
TYPE DFC_MOXEMM_SMU_ALM3_2 : STRUCT
  DTC : UDINT := 16#108900;
  DFCid : UINT := 938;
  debounceMethod : USINT := NATIVE;
END_STRUCT;
END_TYPE

{attribute 'external_name' := 'cmp_rts_DFC_ComCntESP_07'}
TYPE DFC_ComCntESP_07 : STRUCT
  DTC : UDINT := 16#102300;
END_STRUCT;
END_TYPE

{attribute 'external_name' := 'cmp_rts_DFC_MOXEMM_SMU_ALM3_4'}
TYPE DFC_MOXEMM_SMU_ALM3_4 : STRUCT
  DTC : UDINT := 16#108A00;
  DFCid : UINT := 941;
  debounceMethod : USINT := NATIVE;
END_STRUCT;
END_TYPE

{attribute 'external_name' := 'cmp_rts_DFC_MOXEMM_SMU_ALM3_5'}
TYPE DFC_MOXEMM_SMU_ALM3_5 : STRUCT
  DTC : UDINT := 16#108B00;
  DFCid : UINT := 942;
  debounceMethod : USINT := NATIVE;
END_STRUCT;
END_TYPE

{attribute 'external_name' := 'cmp_rts_DFC_MOXEMM_SMU_ALM3_7'}
TYPE DFC_MOXEMM_SMU_ALM3_7 : STRUCT
  DTC : UDINT := 16#108C00;
  DFCid : UINT := 943;
  debounceMethod : USINT := NATIVE;
END_STRUCT;
END_TYPE

{attribute 'external_name' := 'cmp_rts_DFC_MoXEMMHwLTRegMonTest'}
TYPE DFC_MoXEMMHwLTRegMonTest : STRUCT
  DTC : UDINT := 16#10D400;
  DFCid : UINT := 997;
  debounceMethod : USINT := NATIVE;
END_STRUCT;
END_TYPE

{attribute 'external_name' := 'cmp_rts_DFC_ComCntESP_02'}
TYPE DFC_ComCntESP_02 : STRUCT
  DTC : UDINT := 16#102100;
END_STRUCT;
END_TYPE

{attribute 'external_name' := 'cmp_rts_DFC_DSMDummy'}
TYPE DFC_DSMDummy : STRUCT
  DTC : UDINT := 16#100F00;
  DFCid : UINT := 518;
  debounceMethod : USINT := NO_DEBOUNCE;
END_STRUCT;
END_TYPE

{attribute 'external_name' := 'cmp_rts_DFC_MOXEMM_SMU_ALM2_22'}
TYPE DFC_MOXEMM_SMU_ALM2_22 : STRUCT
  DTC : UDINT := 16#108600;
  DFCid : UINT := 927;
  debounceMethod : USINT := NATIVE;
END_STRUCT;
END_TYPE

{attribute 'external_name' := 'cmp_rts_DFC_SWReset'}
TYPE DFC_SWReset : STRUCT
  DTC : UDINT := 16#105600;
  DFCid : UINT := 1004;
  debounceMethod : USINT := NATIVE;
END_STRUCT;
END_TYPE

{attribute 'external_name' := 'cmp_rts_DFC_MOXEMM_SMU_ALM2_23'}
TYPE DFC_MOXEMM_SMU_ALM2_23 : STRUCT
  DTC : UDINT := 16#108700;
  DFCid : UINT := 928;
  debounceMethod : USINT := NATIVE;
END_STRUCT;
END_TYPE

{attribute 'external_name' := 'cmp_rts_DFC_MoXEMMHwLTMBIST'}
TYPE DFC_MoXEMMHwLTMBIST : STRUCT
  DTC : UDINT := 16#10D100;
END_STRUCT;
END_TYPE

{attribute 'external_name' := 'cmp_rts_DFC_MOXEMM_SMU_ALM7_31'}
TYPE DFC_MOXEMM_SMU_ALM7_31 : STRUCT
  DTC : UDINT := 16#10B000;
  DFCid : UINT := 974;
  debounceMethod : USINT := NATIVE;
END_STRUCT;
END_TYPE

{attribute 'external_name' := 'cmp_rts_DFC_MOXEMM_SMU_ALM7_30'}
TYPE DFC_MOXEMM_SMU_ALM7_30 : STRUCT
  DTC : UDINT := 16#10AF00;
  DFCid : UINT := 973;
  debounceMethod : USINT := NATIVE;
END_STRUCT;
END_TYPE

{attribute 'external_name' := 'cmp_rts_DFC_OCWDAErrPin'}
TYPE DFC_OCWDAErrPin : STRUCT
  DTC : UDINT := 16#098B00;
  DFCid : UINT := 1003;
  debounceMethod : USINT := NATIVE;
END_STRUCT;
END_TYPE

{attribute 'external_name' := 'cmp_rts_DFC_ComCntESP_19'}
TYPE DFC_ComCntESP_19 : STRUCT
  DTC : UDINT := 16#102500;
END_STRUCT;
END_TYPE

{attribute 'external_name' := 'cmp_rts_DFC_MOXEMM_SMU_ALM8_10'}
TYPE DFC_MOXEMM_SMU_ALM8_10 : STRUCT
  DTC : UDINT := 16#10B600;
  DFCid : UINT := 977;
  debounceMethod : USINT := NATIVE;
END_STRUCT;
END_TYPE

{attribute 'external_name' := 'cmp_rts_DFC_MRlySCG'}
TYPE DFC_MRlySCG : STRUCT
  DTC : UDINT := 16#104B00;
END_STRUCT;
END_TYPE

{attribute 'external_name' := 'cmp_rts_DFC_MOXEMM_SMU_ALM8_11'}
TYPE DFC_MOXEMM_SMU_ALM8_11 : STRUCT
  DTC : UDINT := 16#10B700;
  DFCid : UINT := 978;
  debounceMethod : USINT := NATIVE;
END_STRUCT;
END_TYPE

{attribute 'external_name' := 'cmp_rts_DFC_MOXEMM_SMU_ALM8_12'}
TYPE DFC_MOXEMM_SMU_ALM8_12 : STRUCT
  DTC : UDINT := 16#10B800;
  DFCid : UINT := 979;
  debounceMethod : USINT := NATIVE;
END_STRUCT;
END_TYPE

{attribute 'external_name' := 'cmp_rts_DFC_MOXEMM_SMU_ALM8_13'}
TYPE DFC_MOXEMM_SMU_ALM8_13 : STRUCT
  DTC : UDINT := 16#10B900;
  DFCid : UINT := 980;
  debounceMethod : USINT := NATIVE;
END_STRUCT;
END_TYPE

{attribute 'external_name' := 'cmp_rts_DFC_MRlySCB'}
TYPE DFC_MRlySCB : STRUCT
  DTC : UDINT := 16#104A00;
END_STRUCT;
END_TYPE

{attribute 'external_name' := 'cmp_rts_DFC_MoXEMMHwLTMCUFW'}
TYPE DFC_MoXEMMHwLTMCUFW : STRUCT
  DTC : UDINT := 16#10D200;
  DFCid : UINT := 995;
  debounceMethod : USINT := NATIVE;
END_STRUCT;
END_TYPE

{attribute 'external_name' := 'cmp_rts_DFC_MOXEMM_SMU_ALM8_16'}
TYPE DFC_MOXEMM_SMU_ALM8_16 : STRUCT
  DTC : UDINT := 16#10BA00;
  DFCid : UINT := 981;
  debounceMethod : USINT := NATIVE;
END_STRUCT;
END_TYPE

{attribute 'external_name' := 'cmp_rts_DFC_MOXEMM_SMU_ALM8_18'}
TYPE DFC_MOXEMM_SMU_ALM8_18 : STRUCT
  DTC : UDINT := 16#10BB00;
  DFCid : UINT := 982;
  debounceMethod : USINT := NATIVE;
END_STRUCT;
END_TYPE

{attribute 'external_name' := 'cmp_rts_DFC_ComCntESP_10'}
TYPE DFC_ComCntESP_10 : STRUCT
  DTC : UDINT := 16#102400;
END_STRUCT;
END_TYPE

{attribute 'external_name' := 'cmp_rts_DFC_CAN_E_TIMEOUT'}
TYPE DFC_CAN_E_TIMEOUT : STRUCT
  DTC : UDINT := 16#094200;
  DFCid : UINT := 861;
  debounceMethod : USINT := NO_DEBOUNCE;
END_STRUCT;
END_TYPE

{attribute 'external_name' := 'cmp_rts_DFC_RBA_IOEXTLIB_KEEPALIVE_INI'}
TYPE DFC_RBA_IOEXTLIB_KEEPALIVE_INI : STRUCT
  DTC : UDINT := 16#094400;
  DFCid : UINT := 872;
  debounceMethod : USINT := NO_DEBOUNCE;
END_STRUCT;
END_TYPE

{attribute 'external_name' := 'cmp_rts_DFC_Com_vWhlRrL'}
TYPE DFC_Com_vWhlRrL : STRUCT
  DTC : UDINT := 16#103D00;
END_STRUCT;
END_TYPE

{attribute 'external_name' := 'cmp_rts_DFC_Com_numWhlIncFrtLeft'}
TYPE DFC_Com_numWhlIncFrtLeft : STRUCT
  DTC : UDINT := 16#103A00;
END_STRUCT;
END_TYPE

{attribute 'external_name' := 'cmp_rts_DFC_rba_MemDiag_MemWrErr'}
TYPE DFC_rba_MemDiag_MemWrErr : STRUCT
  DTC : UDINT := 16#094800;
  DFCid : UINT := 876;
  debounceMethod : USINT := NO_DEBOUNCE;
END_STRUCT;
END_TYPE

{attribute 'external_name' := 'cmp_rts_DFC_CANTRCV_E_NO_TRCV_CONTROL_0'}
TYPE DFC_CANTRCV_E_NO_TRCV_CONTROL_0 : STRUCT
  DTC : UDINT := 16#094000;
  DFCid : UINT := 860;
  debounceMethod : USINT := NO_DEBOUNCE;
END_STRUCT;
END_TYPE

{attribute 'external_name' := 'cmp_rts_DFC_MOXEMM_SMU_ALM3_11'}
TYPE DFC_MOXEMM_SMU_ALM3_11 : STRUCT
  DTC : UDINT := 16#108F00;
  DFCid : UINT := 935;
  debounceMethod : USINT := NATIVE;
END_STRUCT;
END_TYPE

{attribute 'external_name' := 'cmp_rts_DFC_MOXEMM_SMU_ALM3_14'}
TYPE DFC_MOXEMM_SMU_ALM3_14 : STRUCT
  DTC : UDINT := 16#109100;
  DFCid : UINT := 937;
  debounceMethod : USINT := NATIVE;
END_STRUCT;
END_TYPE

{attribute 'external_name' := 'cmp_rts_DFC_MOXEMM_SMU_ALM3_13'}
TYPE DFC_MOXEMM_SMU_ALM3_13 : STRUCT
  DTC : UDINT := 16#109000;
  DFCid : UINT := 936;
  debounceMethod : USINT := NATIVE;
END_STRUCT;
END_TYPE

{attribute 'external_name' := 'cmp_rts_DFC_MOXEMM_SMU_ALM3_10'}
TYPE DFC_MOXEMM_SMU_ALM3_10 : STRUCT
  DTC : UDINT := 16#108E00;
  DFCid : UINT := 934;
  debounceMethod : USINT := NATIVE;
END_STRUCT;
END_TYPE

{attribute 'external_name' := 'cmp_rts_DFC_MOXEMM_SMU_ALM8_30'}
TYPE DFC_MOXEMM_SMU_ALM8_30 : STRUCT
  DTC : UDINT := 16#10BC00;
  DFCid : UINT := 985;
  debounceMethod : USINT := NATIVE;
END_STRUCT;
END_TYPE

{attribute 'external_name' := 'cmp_rts_DFC_MOXEMM_SMU_ALM8_31'}
TYPE DFC_MOXEMM_SMU_ALM8_31 : STRUCT
  DTC : UDINT := 16#10BD00;
  DFCid : UINT := 986;
  debounceMethod : USINT := NATIVE;
END_STRUCT;
END_TYPE

{attribute 'external_name' := 'cmp_rts_DFC_ComCntACC_06'}
TYPE DFC_ComCntACC_06 : STRUCT
  DTC : UDINT := 16#101F00;
END_STRUCT;
END_TYPE

{attribute 'external_name' := 'cmp_rts_DFC_rba_T15_Diag_ComInVld_Event'}
TYPE DFC_rba_T15_Diag_ComInVld_Event : STRUCT
  DTC : UDINT := 16#094B00;
  DFCid : UINT := 878;
  debounceMethod : USINT := NO_DEBOUNCE;
END_STRUCT;
END_TYPE

{attribute 'external_name' := 'cmp_rts_DFC_MOXEMM_SMU_ALM11_0'}
TYPE DFC_MOXEMM_SMU_ALM11_0 : STRUCT
  DTC : UDINT := 16#10C500;
  DFCid : UINT := 897;
  debounceMethod : USINT := NATIVE;
END_STRUCT;
END_TYPE

{attribute 'external_name' := 'cmp_rts_DFC_MOXEMM_SMU_ALM11_1'}
TYPE DFC_MOXEMM_SMU_ALM11_1 : STRUCT
  DTC : UDINT := 16#10C600;
  DFCid : UINT := 898;
  debounceMethod : USINT := NATIVE;
END_STRUCT;
END_TYPE

{attribute 'external_name' := 'cmp_rts_DFC_MOXEMM_SMU_ALM11_2'}
TYPE DFC_MOXEMM_SMU_ALM11_2 : STRUCT
  DTC : UDINT := 16#10C700;
  DFCid : UINT := 899;
  debounceMethod : USINT := NATIVE;
END_STRUCT;
END_TYPE

{attribute 'external_name' := 'cmp_rts_DFC_MOXEMM_SMU_ALM3_23'}
TYPE DFC_MOXEMM_SMU_ALM3_23 : STRUCT
  DTC : UDINT := 16#109300;
  DFCid : UINT := 940;
  debounceMethod : USINT := NATIVE;
END_STRUCT;
END_TYPE

{attribute 'external_name' := 'cmp_rts_DFC_MOXEMM_SMU_ALM3_22'}
TYPE DFC_MOXEMM_SMU_ALM3_22 : STRUCT
  DTC : UDINT := 16#109200;
  DFCid : UINT := 939;
  debounceMethod : USINT := NATIVE;
END_STRUCT;
END_TYPE

{attribute 'external_name' := 'cmp_rts_DFC_OCWDACom'}
TYPE DFC_OCWDACom : STRUCT
  DTC : UDINT := 16#098A00;
  DFCid : UINT := 1002;
  debounceMethod : USINT := NATIVE;
END_STRUCT;
END_TYPE

{attribute 'external_name' := 'cmp_rts_DFC_MoFVarPostBldSel'}
TYPE DFC_MoFVarPostBldSel : STRUCT
  DTC : UDINT := 16#098900;
  DFCid : UINT := 993;
  debounceMethod : USINT := NATIVE;
END_STRUCT;
END_TYPE

{attribute 'external_name' := 'cmp_rts_DFC_MOXEMM_SMU_ALM1_2'}
TYPE DFC_MOXEMM_SMU_ALM1_2 : STRUCT
  DTC : UDINT := 16#107100;
  DFCid : UINT := 911;
  debounceMethod : USINT := NATIVE;
END_STRUCT;
END_TYPE

{attribute 'external_name' := 'cmp_rts_DFC_MOXEMM_SMU_ALM1_4'}
TYPE DFC_MOXEMM_SMU_ALM1_4 : STRUCT
  DTC : UDINT := 16#107200;
  DFCid : UINT := 914;
  debounceMethod : USINT := NATIVE;
END_STRUCT;
END_TYPE

{attribute 'external_name' := 'cmp_rts_DFC_MOXEMM_SMU_ALM1_5'}
TYPE DFC_MOXEMM_SMU_ALM1_5 : STRUCT
  DTC : UDINT := 16#107300;
  DFCid : UINT := 915;
  debounceMethod : USINT := NATIVE;
END_STRUCT;
END_TYPE

{attribute 'external_name' := 'cmp_rts_DFC_MOXEMM_SMU_ALM1_7'}
TYPE DFC_MOXEMM_SMU_ALM1_7 : STRUCT
  DTC : UDINT := 16#107400;
  DFCid : UINT := 916;
  debounceMethod : USINT := NATIVE;
END_STRUCT;
END_TYPE

{attribute 'external_name' := 'cmp_rts_DFC_MOXEMM_SMU_ALM1_8'}
TYPE DFC_MOXEMM_SMU_ALM1_8 : STRUCT
  DTC : UDINT := 16#107500;
  DFCid : UINT := 917;
  debounceMethod : USINT := NATIVE;
END_STRUCT;
END_TYPE

{attribute 'external_name' := 'cmp_rts_DFC_MOXEMM_SMU_ALM9_0'}
TYPE DFC_MOXEMM_SMU_ALM9_0 : STRUCT
  DTC : UDINT := 16#10BE00;
  DFCid : UINT := 988;
  debounceMethod : USINT := NATIVE;
END_STRUCT;
END_TYPE

{attribute 'external_name' := 'cmp_rts_DFC_MOXEMM_SMU_ALM9_1'}
TYPE DFC_MOXEMM_SMU_ALM9_1 : STRUCT
  DTC : UDINT := 16#10BF00;
  DFCid : UINT := 989;
  debounceMethod : USINT := NATIVE;
END_STRUCT;
END_TYPE

{attribute 'external_name' := 'cmp_rts_DFC_ComChksBMS_01'}
TYPE DFC_ComChksBMS_01 : STRUCT
  DTC : UDINT := 16#101700;
END_STRUCT;
END_TYPE

{attribute 'external_name' := 'cmp_rts_DFC_LIN_E_TIMEOUT'}
TYPE DFC_LIN_E_TIMEOUT : STRUCT
  DTC : UDINT := 16#094100;
  DFCid : UINT := 868;
  debounceMethod : USINT := NO_DEBOUNCE;
END_STRUCT;
END_TYPE

{attribute 'external_name' := 'cmp_rts_DFC_MOXEMM_SMU_ALM1_0'}
TYPE DFC_MOXEMM_SMU_ALM1_0 : STRUCT
  DTC : UDINT := 16#106F00;
  DFCid : UINT := 905;
  debounceMethod : USINT := NATIVE;
END_STRUCT;
END_TYPE

{attribute 'external_name' := 'cmp_rts_DFC_MOXEMM_SMU_ALM1_1'}
TYPE DFC_MOXEMM_SMU_ALM1_1 : STRUCT
  DTC : UDINT := 16#107000;
  DFCid : UINT := 906;
  debounceMethod : USINT := NATIVE;
END_STRUCT;
END_TYPE

{attribute 'external_name' := 'cmp_rts_DFC_MOXEMM_SMU_ALM1_14'}
TYPE DFC_MOXEMM_SMU_ALM1_14 : STRUCT
  DTC : UDINT := 16#107900;
  DFCid : UINT := 910;
  debounceMethod : USINT := NATIVE;
END_STRUCT;
END_TYPE

{attribute 'external_name' := 'cmp_rts_DFC_MOXEMM_SMU_ALM1_13'}
TYPE DFC_MOXEMM_SMU_ALM1_13 : STRUCT
  DTC : UDINT := 16#107800;
  DFCid : UINT := 909;
  debounceMethod : USINT := NATIVE;
END_STRUCT;
END_TYPE

{attribute 'external_name' := 'cmp_rts_DFC_MOXEMM_SMU_ALM1_10'}
TYPE DFC_MOXEMM_SMU_ALM1_10 : STRUCT
  DTC : UDINT := 16#107600;
  DFCid : UINT := 907;
  debounceMethod : USINT := NATIVE;
END_STRUCT;
END_TYPE

{attribute 'external_name' := 'cmp_rts_DFC_rba_T15_Diag_ComOff_HwOn_Event'}
TYPE DFC_rba_T15_Diag_ComOff_HwOn_Event : STRUCT
  DTC : UDINT := 16#094C00;
  DFCid : UINT := 879;
  debounceMethod : USINT := NO_DEBOUNCE;
END_STRUCT;
END_TYPE

{attribute 'external_name' := 'cmp_rts_DFC_MOXEMM_SMU_ALM1_11'}
TYPE DFC_MOXEMM_SMU_ALM1_11 : STRUCT
  DTC : UDINT := 16#107700;
  DFCid : UINT := 908;
  debounceMethod : USINT := NATIVE;
END_STRUCT;
END_TYPE

{attribute 'external_name' := 'cmp_rts_DFC_MOXEMM_SMU_ALM6_25'}
TYPE DFC_MOXEMM_SMU_ALM6_25 : STRUCT
  DTC : UDINT := 16#10A100;
  DFCid : UINT := 955;
  debounceMethod : USINT := NATIVE;
END_STRUCT;
END_TYPE

{attribute 'external_name' := 'cmp_rts_DFC_MOXEMM_SMU_ALM6_21'}
TYPE DFC_MOXEMM_SMU_ALM6_21 : STRUCT
  DTC : UDINT := 16#10A000;
  DFCid : UINT := 954;
  debounceMethod : USINT := NATIVE;
END_STRUCT;
END_TYPE

{attribute 'external_name' := 'cmp_rts_DFC_MOXEMM_SMU_ALM6_20'}
TYPE DFC_MOXEMM_SMU_ALM6_20 : STRUCT
  DTC : UDINT := 16#109F00;
  DFCid : UINT := 953;
  debounceMethod : USINT := NATIVE;
END_STRUCT;
END_TYPE

{attribute 'external_name' := 'cmp_rts_DFC_ComDlcESP_02'}
TYPE DFC_ComDlcESP_02 : STRUCT
  DTC : UDINT := 16#102900;
END_STRUCT;
END_TYPE

{attribute 'external_name' := 'cmp_rts_DFC_MOXEMM_SMU_ALM1_23'}
TYPE DFC_MOXEMM_SMU_ALM1_23 : STRUCT
  DTC : UDINT := 16#107B00;
  DFCid : UINT := 913;
  debounceMethod : USINT := NATIVE;
END_STRUCT;
END_TYPE

{attribute 'external_name' := 'cmp_rts_DFC_MOXEMM_SMU_ALM1_22'}
TYPE DFC_MOXEMM_SMU_ALM1_22 : STRUCT
  DTC : UDINT := 16#107A00;
  DFCid : UINT := 912;
  debounceMethod : USINT := NATIVE;
END_STRUCT;
END_TYPE

{attribute 'external_name' := 'cmp_rts_DFC_rba_MRly_Diag_Stk_Event'}
TYPE DFC_rba_MRly_Diag_Stk_Event : STRUCT
  DTC : UDINT := 16#094600;
  DFCid : UINT := 873;
  debounceMethod : USINT := NO_DEBOUNCE;
END_STRUCT;
END_TYPE

{attribute 'external_name' := 'cmp_rts_DFC_ComDlcESP_05'}
TYPE DFC_ComDlcESP_05 : STRUCT
  DTC : UDINT := 16#102A00;
END_STRUCT;
END_TYPE

{attribute 'external_name' := 'cmp_rts_DFC_DevLibBattULo'}
TYPE DFC_DevLibBattULo : STRUCT
  DTC : UDINT := 16#092400;
  DFCid : UINT := 4;
  debounceMethod : USINT := TIME_UP_DOWN;
END_STRUCT;
END_TYPE

{attribute 'external_name' := 'cmp_rts_DFC_ComDlcESP_07'}
TYPE DFC_ComDlcESP_07 : STRUCT
  DTC : UDINT := 16#102B00;
END_STRUCT;
END_TYPE

{attribute 'external_name' := 'cmp_rts_DFC_MOXEMM_SMU_ALM2_1'}
TYPE DFC_MOXEMM_SMU_ALM2_1 : STRUCT
  DTC : UDINT := 16#107C00;
  DFCid : UINT := 921;
  debounceMethod : USINT := NATIVE;
END_STRUCT;
END_TYPE

{attribute 'external_name' := 'cmp_rts_DFC_MOXEMM_SMU_ALM2_2'}
TYPE DFC_MOXEMM_SMU_ALM2_2 : STRUCT
  DTC : UDINT := 16#107D00;
  DFCid : UINT := 926;
  debounceMethod : USINT := NATIVE;
END_STRUCT;
END_TYPE

{attribute 'external_name' := 'cmp_rts_DFC_MOXEMM_SMU_ALM2_4'}
TYPE DFC_MOXEMM_SMU_ALM2_4 : STRUCT
  DTC : UDINT := 16#107E00;
  DFCid : UINT := 929;
  debounceMethod : USINT := NATIVE;
END_STRUCT;
END_TYPE

{attribute 'external_name' := 'cmp_rts_DFC_MOXEMM_SMU_ALM2_5'}
TYPE DFC_MOXEMM_SMU_ALM2_5 : STRUCT
  DTC : UDINT := 16#107F00;
  DFCid : UINT := 930;
  debounceMethod : USINT := NATIVE;
END_STRUCT;
END_TYPE

{attribute 'external_name' := 'cmp_rts_DFC_MOXEMM_SMU_ALM2_7'}
TYPE DFC_MOXEMM_SMU_ALM2_7 : STRUCT
  DTC : UDINT := 16#108000;
  DFCid : UINT := 931;
  debounceMethod : USINT := NATIVE;
END_STRUCT;
END_TYPE

{attribute 'external_name' := 'cmp_rts_DFC_MOXEMM_SMU_ALM2_8'}
TYPE DFC_MOXEMM_SMU_ALM2_8 : STRUCT
  DTC : UDINT := 16#108100;
  DFCid : UINT := 932;
  debounceMethod : USINT := NATIVE;
END_STRUCT;
END_TYPE

{attribute 'external_name' := 'cmp_rts_DFC_rba_SyC_IrrSwOffTrigEngRun_Event'}
TYPE DFC_rba_SyC_IrrSwOffTrigEngRun_Event : STRUCT
  DTC : UDINT := 16#094A00;
  DFCid : UINT := 877;
  debounceMethod : USINT := NO_DEBOUNCE;
END_STRUCT;
END_TYPE

{attribute 'external_name' := 'cmp_rts_DFC_ComDlcESP_10'}
TYPE DFC_ComDlcESP_10 : STRUCT
  DTC : UDINT := 16#102C00;
END_STRUCT;
END_TYPE

{attribute 'external_name' := 'cmp_rts_DFC_MOXEMM_SMU_ALM7_17'}
TYPE DFC_MOXEMM_SMU_ALM7_17 : STRUCT
  DTC : UDINT := 16#10A900;
  DFCid : UINT := 966;
  debounceMethod : USINT := NATIVE;
END_STRUCT;
END_TYPE

{attribute 'external_name' := 'cmp_rts_DFC_MOXEMM_SMU_ALM7_16'}
TYPE DFC_MOXEMM_SMU_ALM7_16 : STRUCT
  DTC : UDINT := 16#10A800;
  DFCid : UINT := 965;
  debounceMethod : USINT := NATIVE;
END_STRUCT;
END_TYPE

{attribute 'external_name' := 'cmp_rts_DFC_MOXEMM_SMU_ALM7_15'}
TYPE DFC_MOXEMM_SMU_ALM7_15 : STRUCT
  DTC : UDINT := 16#10A700;
  DFCid : UINT := 964;
  debounceMethod : USINT := NATIVE;
END_STRUCT;
END_TYPE

{attribute 'external_name' := 'cmp_rts_DFC_MOXEMM_SMU_ALM7_14'}
TYPE DFC_MOXEMM_SMU_ALM7_14 : STRUCT
  DTC : UDINT := 16#10A600;
  DFCid : UINT := 963;
  debounceMethod : USINT := NATIVE;
END_STRUCT;
END_TYPE

{attribute 'external_name' := 'cmp_rts_DFC_MOXEMM_SMU_ALM7_13'}
TYPE DFC_MOXEMM_SMU_ALM7_13 : STRUCT
  DTC : UDINT := 16#10A500;
  DFCid : UINT := 962;
  debounceMethod : USINT := NATIVE;
END_STRUCT;
END_TYPE

{attribute 'external_name' := 'cmp_rts_DFC_MOXEMM_SMU_ALM7_12'}
TYPE DFC_MOXEMM_SMU_ALM7_12 : STRUCT
  DTC : UDINT := 16#10A400;
  DFCid : UINT := 961;
  debounceMethod : USINT := NATIVE;
END_STRUCT;
END_TYPE

{attribute 'external_name' := 'cmp_rts_DFC_ComDlcESP_19'}
TYPE DFC_ComDlcESP_19 : STRUCT
  DTC : UDINT := 16#102D00;
END_STRUCT;
END_TYPE

{attribute 'external_name' := 'cmp_rts_DFC_ComCntKlemmen_Status_01'}
TYPE DFC_ComCntKlemmen_Status_01 : STRUCT
  DTC : UDINT := 16#103900;
END_STRUCT;
END_TYPE

{attribute 'external_name' := 'cmp_rts_DFC_rba_T15_Diag_ComOn_HwOff_Event'}
TYPE DFC_rba_T15_Diag_ComOn_HwOff_Event : STRUCT
  DTC : UDINT := 16#094D00;
  DFCid : UINT := 880;
  debounceMethod : USINT := NO_DEBOUNCE;
END_STRUCT;
END_TYPE

{attribute 'external_name' := 'cmp_rts_DFC_MoXEMMHwLTStbySMUAlvTest'}
TYPE DFC_MoXEMMHwLTStbySMUAlvTest : STRUCT
  DTC : UDINT := 16#10D500;
  DFCid : UINT := 998;
  debounceMethod : USINT := NATIVE;
END_STRUCT;
END_TYPE

{attribute 'external_name' := 'cmp_rts_DFC_rba_MultiStackTrace_Threshold'}
TYPE DFC_rba_MultiStackTrace_Threshold : STRUCT
  DTC : UDINT := 16#094900;
  DFCid : UINT := 869;
  debounceMethod : USINT := NO_DEBOUNCE;
END_STRUCT;
END_TYPE

{attribute 'external_name' := 'cmp_rts_DFC_MOXEMM_SMU_ALM2_14'}
TYPE DFC_MOXEMM_SMU_ALM2_14 : STRUCT
  DTC : UDINT := 16#108500;
  DFCid : UINT := 925;
  debounceMethod : USINT := NATIVE;
END_STRUCT;
END_TYPE

{attribute 'external_name' := 'cmp_rts_DFC_ComDlcESP_20'}
TYPE DFC_ComDlcESP_20 : STRUCT
  DTC : UDINT := 16#102E00;
END_STRUCT;
END_TYPE

{attribute 'external_name' := 'cmp_rts_DFC_MOXEMM_SMU_ALM2_11'}
TYPE DFC_MOXEMM_SMU_ALM2_11 : STRUCT
  DTC : UDINT := 16#108300;
  DFCid : UINT := 923;
  debounceMethod : USINT := NATIVE;
END_STRUCT;
END_TYPE

{attribute 'external_name' := 'cmp_rts_DFC_MOXEMM_SMU_ALM7_29'}
TYPE DFC_MOXEMM_SMU_ALM7_29 : STRUCT
  DTC : UDINT := 16#10AE00;
  DFCid : UINT := 972;
  debounceMethod : USINT := NATIVE;
END_STRUCT;
END_TYPE

{attribute 'external_name' := 'cmp_rts_DFC_ComDlcESP_21'}
TYPE DFC_ComDlcESP_21 : STRUCT
  DTC : UDINT := 16#102F00;
END_STRUCT;
END_TYPE

{attribute 'external_name' := 'cmp_rts_DFC_MOXEMM_SMU_ALM2_10'}
TYPE DFC_MOXEMM_SMU_ALM2_10 : STRUCT
  DTC : UDINT := 16#108200;
  DFCid : UINT := 922;
  debounceMethod : USINT := NATIVE;
END_STRUCT;
END_TYPE

{attribute 'external_name' := 'cmp_rts_DFC_MOXEMM_SMU_ALM7_28'}
TYPE DFC_MOXEMM_SMU_ALM7_28 : STRUCT
  DTC : UDINT := 16#10AD00;
  DFCid : UINT := 971;
  debounceMethod : USINT := NATIVE;
END_STRUCT;
END_TYPE

{attribute 'external_name' := 'cmp_rts_DFC_MOXEMM_SMU_ALM2_13'}
TYPE DFC_MOXEMM_SMU_ALM2_13 : STRUCT
  DTC : UDINT := 16#108400;
  DFCid : UINT := 924;
  debounceMethod : USINT := NATIVE;
END_STRUCT;
END_TYPE

{attribute 'external_name' := 'cmp_rts_DFC_MOXEMM_SMU_ALM7_26'}
TYPE DFC_MOXEMM_SMU_ALM7_26 : STRUCT
  DTC : UDINT := 16#10AC00;
  DFCid : UINT := 970;
  debounceMethod : USINT := NATIVE;
END_STRUCT;
END_TYPE

{attribute 'external_name' := 'cmp_rts_DFC_MOXEMM_SMU_ALM3_8'}
TYPE DFC_MOXEMM_SMU_ALM3_8 : STRUCT
  DTC : UDINT := 16#108D00;
  DFCid : UINT := 944;
  debounceMethod : USINT := NATIVE;
END_STRUCT;
END_TYPE

{attribute 'external_name' := 'cmp_rts_DFC_MOXEMM_SMU_ALM7_25'}
TYPE DFC_MOXEMM_SMU_ALM7_25 : STRUCT
  DTC : UDINT := 16#10AB00;
  DFCid : UINT := 969;
  debounceMethod : USINT := NATIVE;
END_STRUCT;
END_TYPE

{attribute 'external_name' := 'cmp_rts_DFC_MOXEMM_SMU_ALM7_20'}
TYPE DFC_MOXEMM_SMU_ALM7_20 : STRUCT
  DTC : UDINT := 16#10AA00;
  DFCid : UINT := 968;
  debounceMethod : USINT := NATIVE;
END_STRUCT;
END_TYPE

{attribute 'external_name' := 'cmp_rts_DFC_MRlyOL'}
TYPE DFC_MRlyOL : STRUCT
  DTC : UDINT := 16#104900;
END_STRUCT;
END_TYPE

{attribute 'external_name' := 'cmp_rts_DFC_MOXEMM_SMU_ALM7_1'}
TYPE DFC_MOXEMM_SMU_ALM7_1 : STRUCT
  DTC : UDINT := 16#10A200;
  DFCid : UINT := 960;
  debounceMethod : USINT := NATIVE;
END_STRUCT;
END_TYPE

{attribute 'external_name' := 'cmp_rts_DFC_ComChksESP_19'}
TYPE DFC_ComChksESP_19 : STRUCT
  DTC : UDINT := 16#101C00;
END_STRUCT;
END_TYPE

{attribute 'external_name' := 'cmp_rts_DFC_MOXEMM_SMU_ALM7_2'}
TYPE DFC_MOXEMM_SMU_ALM7_2 : STRUCT
  DTC : UDINT := 16#10A300;
  DFCid : UINT := 967;
  debounceMethod : USINT := NATIVE;
END_STRUCT;
END_TYPE

{attribute 'external_name' := 'cmp_rts_DFC_ComTOutESP_10'}
TYPE DFC_ComTOutESP_10 : STRUCT
  DTC : UDINT := 16#103400;
END_STRUCT;
END_TYPE

{attribute 'external_name' := 'cmp_rts_DFC_Com_stWhlSensRrRht'}
TYPE DFC_Com_stWhlSensRrRht : STRUCT
  DTC : UDINT := 16#103B00;
END_STRUCT;
END_TYPE

{attribute 'external_name' := 'cmp_rts_DFC_ComChksKlemmen_Status_01'}
TYPE DFC_ComChksKlemmen_Status_01 : STRUCT
  DTC : UDINT := 16#103800;
END_STRUCT;
END_TYPE

{attribute 'external_name' := 'cmp_rts_DFC_ComTOutESP_07'}
TYPE DFC_ComTOutESP_07 : STRUCT
  DTC : UDINT := 16#103300;
END_STRUCT;
END_TYPE

{attribute 'external_name' := 'cmp_rts_DFC_ComDlcACC_06'}
TYPE DFC_ComDlcACC_06 : STRUCT
  DTC : UDINT := 16#102800;
END_STRUCT;
END_TYPE

{attribute 'external_name' := 'cmp_rts_DFC_rba_MemDiag_MemReadErr'}
TYPE DFC_rba_MemDiag_MemReadErr : STRUCT
  DTC : UDINT := 16#094700;
  DFCid : UINT := 875;
  debounceMethod : USINT := NO_DEBOUNCE;
END_STRUCT;
END_TYPE

{attribute 'external_name' := 'cmp_rts_DFC_ComChksESP_10'}
TYPE DFC_ComChksESP_10 : STRUCT
  DTC : UDINT := 16#101B00;
END_STRUCT;
END_TYPE

{attribute 'external_name' := 'cmp_rts_DFC_ComChksESP_05'}
TYPE DFC_ComChksESP_05 : STRUCT
  DTC : UDINT := 16#101900;
END_STRUCT;
END_TYPE

{attribute 'external_name' := 'cmp_rts_DFC_OCWDAABEActv'}
TYPE DFC_OCWDAABEActv : STRUCT
  DTC : UDINT := 16#10D800;
  DFCid : UINT := 1001;
  debounceMethod : USINT := NATIVE;
END_STRUCT;
END_TYPE

{attribute 'external_name' := 'cmp_rts_DFC_ComChksESP_07'}
TYPE DFC_ComChksESP_07 : STRUCT
  DTC : UDINT := 16#101A00;
END_STRUCT;
END_TYPE

{attribute 'external_name' := 'cmp_rts_DFC_ComTOutESP_21'}
TYPE DFC_ComTOutESP_21 : STRUCT
  DTC : UDINT := 16#103700;
END_STRUCT;
END_TYPE

{attribute 'external_name' := 'cmp_rts_DFC_ComTOutESP_20'}
TYPE DFC_ComTOutESP_20 : STRUCT
  DTC : UDINT := 16#103600;
END_STRUCT;
END_TYPE

{attribute 'external_name' := 'cmp_rts_DFC_MOXEMM_SMU_ALM0_13'}
TYPE DFC_MOXEMM_SMU_ALM0_13 : STRUCT
  DTC : UDINT := 16#106B00;
  DFCid : UINT := 885;
  debounceMethod : USINT := NATIVE;
END_STRUCT;
END_TYPE

{attribute 'external_name' := 'cmp_rts_DFC_MOXEMM_SMU_ALM0_14'}
TYPE DFC_MOXEMM_SMU_ALM0_14 : STRUCT
  DTC : UDINT := 16#106C00;
  DFCid : UINT := 886;
  debounceMethod : USINT := NATIVE;
END_STRUCT;
END_TYPE

{attribute 'external_name' := 'cmp_rts_DFC_ComTOutESP_19'}
TYPE DFC_ComTOutESP_19 : STRUCT
  DTC : UDINT := 16#103500;
END_STRUCT;
END_TYPE

{attribute 'external_name' := 'cmp_rts_DFC_MOXEMM_SMU_ALM0_10'}
TYPE DFC_MOXEMM_SMU_ALM0_10 : STRUCT
  DTC : UDINT := 16#106900;
  DFCid : UINT := 883;
  debounceMethod : USINT := NATIVE;
END_STRUCT;
END_TYPE

{attribute 'external_name' := 'cmp_rts_DFC_MOXEMM_SMU_ALM0_11'}
TYPE DFC_MOXEMM_SMU_ALM0_11 : STRUCT
  DTC : UDINT := 16#106A00;
  DFCid : UINT := 884;
  debounceMethod : USINT := NATIVE;
END_STRUCT;
END_TYPE

{attribute 'external_name' := 'cmp_rts_DFC_MOXEMM_SMU_ALM8_3'}
TYPE DFC_MOXEMM_SMU_ALM8_3 : STRUCT
  DTC : UDINT := 16#10B400;
  DFCid : UINT := 984;
  debounceMethod : USINT := NATIVE;
END_STRUCT;
END_TYPE

{attribute 'external_name' := 'cmp_rts_DFC_MOXEMM_SMU_ALM8_4'}
TYPE DFC_MOXEMM_SMU_ALM8_4 : STRUCT
  DTC : UDINT := 16#10B500;
  DFCid : UINT := 987;
  debounceMethod : USINT := NATIVE;
END_STRUCT;
END_TYPE

{attribute 'external_name' := 'cmp_rts_DFC_ComChksESP_02'}
TYPE DFC_ComChksESP_02 : STRUCT
  DTC : UDINT := 16#101800;
END_STRUCT;
END_TYPE

{attribute 'external_name' := 'cmp_rts_DFC_DevLibBattUHi'}
TYPE DFC_DevLibBattUHi : STRUCT
  DTC : UDINT := 16#092300;
  DFCid : UINT := 3;
  debounceMethod : USINT := TIME_UP_DOWN;
END_STRUCT;
END_TYPE

{attribute 'external_name' := 'cmp_rts_DFC_Com_trqClthTCSDCSDes'}
TYPE DFC_Com_trqClthTCSDCSDes : STRUCT
  DTC : UDINT := 16#103C00;
END_STRUCT;
END_TYPE

{attribute 'external_name' := 'cmp_rts_DFC_MOXEMM_SMU_ALM0_4'}
TYPE DFC_MOXEMM_SMU_ALM0_4 : STRUCT
  DTC : UDINT := 16#106500;
  DFCid : UINT := 890;
  debounceMethod : USINT := NATIVE;
END_STRUCT;
END_TYPE

{attribute 'external_name' := 'cmp_rts_DFC_MoXEMMHwLTTempSens'}
TYPE DFC_MoXEMMHwLTTempSens : STRUCT
  DTC : UDINT := 16#10D600;
  DFCid : UINT := 999;
  debounceMethod : USINT := NATIVE;
END_STRUCT;
END_TYPE

{attribute 'external_name' := 'cmp_rts_DFC_MOXEMM_SMU_ALM0_5'}
TYPE DFC_MOXEMM_SMU_ALM0_5 : STRUCT
  DTC : UDINT := 16#106600;
  DFCid : UINT := 891;
  debounceMethod : USINT := NATIVE;
END_STRUCT;
END_TYPE

{attribute 'external_name' := 'cmp_rts_DFC_MOXEMM_SMU_ALM0_7'}
TYPE DFC_MOXEMM_SMU_ALM0_7 : STRUCT
  DTC : UDINT := 16#106700;
  DFCid : UINT := 892;
  debounceMethod : USINT := NATIVE;
END_STRUCT;
END_TYPE

{attribute 'external_name' := 'cmp_rts_DFC_MOXEMM_SMU_ALM0_8'}
TYPE DFC_MOXEMM_SMU_ALM0_8 : STRUCT
  DTC : UDINT := 16#106800;
  DFCid : UINT := 893;
  debounceMethod : USINT := NATIVE;
END_STRUCT;
END_TYPE

{attribute 'external_name' := 'cmp_rts_DFC_MOXEMM_SMU_ALM8_0'}
TYPE DFC_MOXEMM_SMU_ALM8_0 : STRUCT
  DTC : UDINT := 16#10B100;
  DFCid : UINT := 975;
  debounceMethod : USINT := NATIVE;
END_STRUCT;
END_TYPE

{attribute 'external_name' := 'cmp_rts_DFC_MOXEMM_SMU_ALM8_1'}
TYPE DFC_MOXEMM_SMU_ALM8_1 : STRUCT
  DTC : UDINT := 16#10B200;
  DFCid : UINT := 976;
  debounceMethod : USINT := NATIVE;
END_STRUCT;
END_TYPE

{attribute 'external_name' := 'cmp_rts_DFC_MOXEMM_SMU_ALM8_2'}
TYPE DFC_MOXEMM_SMU_ALM8_2 : STRUCT
  DTC : UDINT := 16#10B300;
  DFCid : UINT := 983;
  debounceMethod : USINT := NATIVE;
END_STRUCT;
END_TYPE

{attribute 'external_name' := 'cmp_rts_DFC_ComChksACC_06'}
TYPE DFC_ComChksACC_06 : STRUCT
  DTC : UDINT := 16#101600;
END_STRUCT;
END_TYPE

{attribute 'external_name' := 'cmp_rts_DFC_MOXEMM_SMU_ALM0_0'}
TYPE DFC_MOXEMM_SMU_ALM0_0 : STRUCT
  DTC : UDINT := 16#106200;
  DFCid : UINT := 881;
  debounceMethod : USINT := NATIVE;
END_STRUCT;
END_TYPE

{attribute 'external_name' := 'cmp_rts_DFC_MOXEMM_SMU_ALM0_1'}
TYPE DFC_MOXEMM_SMU_ALM0_1 : STRUCT
  DTC : UDINT := 16#106300;
  DFCid : UINT := 882;
  debounceMethod : USINT := NATIVE;
END_STRUCT;
END_TYPE

{attribute 'external_name' := 'cmp_rts_DFC_SWReset_2'}
TYPE DFC_SWReset_2 : STRUCT
  DTC : UDINT := 16#105900;
END_STRUCT;
END_TYPE

{attribute 'external_name' := 'cmp_rts_DFC_MOXEMM_SMU_ALM0_2'}
TYPE DFC_MOXEMM_SMU_ALM0_2 : STRUCT
  DTC : UDINT := 16#106400;
  DFCid : UINT := 887;
  debounceMethod : USINT := NATIVE;
END_STRUCT;
END_TYPE

{attribute 'external_name' := 'cmp_rts_DFC_MOXEMM_SMU_ALM0_23'}
TYPE DFC_MOXEMM_SMU_ALM0_23 : STRUCT
  DTC : UDINT := 16#106E00;
  DFCid : UINT := 889;
  debounceMethod : USINT := NATIVE;
END_STRUCT;
END_TYPE

{attribute 'external_name' := 'cmp_rts_DFC_MOXEMM_SMU_ALM0_22'}
TYPE DFC_MOXEMM_SMU_ALM0_22 : STRUCT
  DTC : UDINT := 16#106D00;
  DFCid : UINT := 888;
  debounceMethod : USINT := NATIVE;
END_STRUCT;
END_TYPE

{attribute 'external_name' := 'cmp_rts_DFC_ComTOutESP_05'}
TYPE DFC_ComTOutESP_05 : STRUCT
  DTC : UDINT := 16#103200;
END_STRUCT;
END_TYPE

{attribute 'external_name' := 'cmp_rts_DFC_ComTOutESP_02'}
TYPE DFC_ComTOutESP_02 : STRUCT
  DTC : UDINT := 16#103100;
END_STRUCT;
END_TYPE

{attribute 'external_name' := 'cmp_rts_DFC_MOXEMM_SMU_ALM6_18'}
TYPE DFC_MOXEMM_SMU_ALM6_18 : STRUCT
  DTC : UDINT := 16#109E00;
  DFCid : UINT := 951;
  debounceMethod : USINT := NATIVE;
END_STRUCT;
END_TYPE

{attribute 'external_name' := 'cmp_rts_DFC_MOXEMM_SMU_ALM6_17'}
TYPE DFC_MOXEMM_SMU_ALM6_17 : STRUCT
  DTC : UDINT := 16#109D00;
  DFCid : UINT := 950;
  debounceMethod : USINT := NATIVE;
END_STRUCT;
END_TYPE

{attribute 'external_name' := 'cmp_rts_DFC_MOXEMM_SMU_ALM6_15'}
TYPE DFC_MOXEMM_SMU_ALM6_15 : STRUCT
  DTC : UDINT := 16#109C00;
  DFCid : UINT := 949;
  debounceMethod : USINT := NATIVE;
END_STRUCT;
END_TYPE

{attribute 'external_name' := 'cmp_rts_DFC_MOXEMM_SMU_ALM21_16'}
TYPE DFC_MOXEMM_SMU_ALM21_16 : STRUCT
  DTC : UDINT := 16#10CF00;
  DFCid : UINT := 919;
  debounceMethod : USINT := NATIVE;
END_STRUCT;
END_TYPE

{attribute 'external_name' := 'cmp_rts_DFC_MOXEMM_SMU_ALM6_14'}
TYPE DFC_MOXEMM_SMU_ALM6_14 : STRUCT
  DTC : UDINT := 16#109B00;
  DFCid : UINT := 948;
  debounceMethod : USINT := NATIVE;
END_STRUCT;
END_TYPE

{attribute 'external_name' := 'cmp_rts_DFC_MOXEMM_SMU_ALM6_12'}
TYPE DFC_MOXEMM_SMU_ALM6_12 : STRUCT
  DTC : UDINT := 16#109A00;
  DFCid : UINT := 947;
  debounceMethod : USINT := NATIVE;
END_STRUCT;
END_TYPE

{attribute 'external_name' := 'cmp_rts_DFC_MOXEMM_SMU_ALM9_3'}
TYPE DFC_MOXEMM_SMU_ALM9_3 : STRUCT
  DTC : UDINT := 16#10C000;
  DFCid : UINT := 991;
  debounceMethod : USINT := NATIVE;
END_STRUCT;
END_TYPE

{attribute 'external_name' := 'cmp_rts_DFC_MOXEMM_SMU_ALM6_11'}
TYPE DFC_MOXEMM_SMU_ALM6_11 : STRUCT
  DTC : UDINT := 16#109900;
  DFCid : UINT := 946;
  debounceMethod : USINT := NATIVE;
END_STRUCT;
END_TYPE

{attribute 'external_name' := 'cmp_rts_DFC_ComTOutACC_06'}
TYPE DFC_ComTOutACC_06 : STRUCT
  DTC : UDINT := 16#103000;
END_STRUCT;
END_TYPE

{attribute 'external_name' := 'cmp_rts_DFC_MOXEMM_SMU_ALM9_15'}
TYPE DFC_MOXEMM_SMU_ALM9_15 : STRUCT
  DTC : UDINT := 16#10C100;
  DFCid : UINT := 990;
  debounceMethod : USINT := NATIVE;
END_STRUCT;
END_TYPE

{attribute 'external_name' := 'cmp_rts_DFC_MOXEMM_SMU_ALM11_8'}
TYPE DFC_MOXEMM_SMU_ALM11_8 : STRUCT
  DTC : UDINT := 16#10CB00;
  DFCid : UINT := 903;
  debounceMethod : USINT := NATIVE;
END_STRUCT;
END_TYPE

{attribute 'external_name' := 'cmp_rts_DFC_MOXEMM_SMU_ALM11_9'}
TYPE DFC_MOXEMM_SMU_ALM11_9 : STRUCT
  DTC : UDINT := 16#10CC00;
  DFCid : UINT := 904;
  debounceMethod : USINT := NATIVE;
END_STRUCT;
END_TYPE

{attribute 'external_name' := 'cmp_rts_DFC_MOXEMM_SMU_ALM11_3'}
TYPE DFC_MOXEMM_SMU_ALM11_3 : STRUCT
  DTC : UDINT := 16#10C800;
  DFCid : UINT := 900;
  debounceMethod : USINT := NATIVE;
END_STRUCT;
END_TYPE

{attribute 'external_name' := 'cmp_rts_DFC_MOXEMM_SMU_ALM11_4'}
TYPE DFC_MOXEMM_SMU_ALM11_4 : STRUCT
  DTC : UDINT := 16#10C900;
  DFCid : UINT := 901;
  debounceMethod : USINT := NATIVE;
END_STRUCT;
END_TYPE

{attribute 'external_name' := 'cmp_rts_DFC_MOXEMM_SMU_ALM11_5'}
TYPE DFC_MOXEMM_SMU_ALM11_5 : STRUCT
  DTC : UDINT := 16#10CA00;
  DFCid : UINT := 902;
  debounceMethod : USINT := NATIVE;
END_STRUCT;
END_TYPE

{attribute 'external_name' := 'cmp_rts_DFC_MOXEMM_SMU_ALM10_16'}
TYPE DFC_MOXEMM_SMU_ALM10_16 : STRUCT
  DTC : UDINT := 16#10C200;
  DFCid : UINT := 894;
  debounceMethod : USINT := NATIVE;
END_STRUCT;
END_TYPE

{attribute 'external_name' := 'cmp_rts_DFC_MOXEMM_SMU_ALM10_17'}
TYPE DFC_MOXEMM_SMU_ALM10_17 : STRUCT
  DTC : UDINT := 16#10C300;
  DFCid : UINT := 895;
  debounceMethod : USINT := NATIVE;
END_STRUCT;
END_TYPE

{attribute 'external_name' := 'cmp_rts_DFC_MoXEMMHwLTUCBCfg'}
TYPE DFC_MoXEMMHwLTUCBCfg : STRUCT
  DTC : UDINT := 16#10D700;
  DFCid : UINT := 1000;
  debounceMethod : USINT := NATIVE;
END_STRUCT;
END_TYPE

{attribute 'external_name' := 'cmp_rts_DFC_CANSM_E_BUS_OFF_NETWORK_0'}
TYPE DFC_CANSM_E_BUS_OFF_NETWORK_0 : STRUCT
  DTC : UDINT := 16#104C00;
  DFCid : UINT := 856;
  debounceMethod : USINT := NO_DEBOUNCE;
END_STRUCT;
END_TYPE

{attribute 'external_name' := 'cmp_rts_DFC_CANSM_E_BUS_OFF_NETWORK_3'}
TYPE DFC_CANSM_E_BUS_OFF_NETWORK_3 : STRUCT
  DTC : UDINT := 16#104F00;
  DFCid : UINT := 859;
  debounceMethod : USINT := NO_DEBOUNCE;
END_STRUCT;
END_TYPE

{attribute 'external_name' := 'cmp_rts_DFC_CANSM_E_BUS_OFF_NETWORK_1'}
TYPE DFC_CANSM_E_BUS_OFF_NETWORK_1 : STRUCT
  DTC : UDINT := 16#104D00;
  DFCid : UINT := 857;
  debounceMethod : USINT := NO_DEBOUNCE;
END_STRUCT;
END_TYPE

{attribute 'external_name' := 'cmp_rts_DFC_CANSM_E_BUS_OFF_NETWORK_2'}
TYPE DFC_CANSM_E_BUS_OFF_NETWORK_2 : STRUCT
  DTC : UDINT := 16#104E00;
  DFCid : UINT := 858;
  debounceMethod : USINT := NO_DEBOUNCE;
END_STRUCT;
END_TYPE

{attribute 'external_name' := 'cmp_rts_DFC_ComCntBMS_01'}
TYPE DFC_ComCntBMS_01 : STRUCT
  DTC : UDINT := 16#102000;
END_STRUCT;
END_TYPE

{attribute 'external_name' := 'cmp_rts_DFC_MoXEMMHwLTLBIST'}
TYPE DFC_MoXEMMHwLTLBIST : STRUCT
  DTC : UDINT := 16#10D000;
END_STRUCT;
END_TYPE

{attribute 'external_name' := 'cmp_rts_DFC_MoXEMMHwLTMonBIST'}
TYPE DFC_MoXEMMHwLTMonBIST : STRUCT
  DTC : UDINT := 16#10D300;
  DFCid : UINT := 996;
  debounceMethod : USINT := NATIVE;
END_STRUCT;
END_TYPE

{attribute 'external_name' := 'cmp_rts_DFC_SWReset_1'}
TYPE DFC_SWReset_1 : STRUCT
  DTC : UDINT := 16#105800;
END_STRUCT;
END_TYPE

{attribute 'external_name' := 'cmp_rts_DFC_SWReset_0'}
TYPE DFC_SWReset_0 : STRUCT
  DTC : UDINT := 16#105700;
END_STRUCT;
END_TYPE

{attribute 'external_name' := 'cmp_rts_DFC_rba_MemDiagExtd_MemReadSngErr'}
TYPE DFC_rba_MemDiagExtd_MemReadSngErr : STRUCT
  DTC : UDINT := 16#103E00;
  DFCid : UINT := 874;
  debounceMethod : USINT := NO_DEBOUNCE;
END_STRUCT;
END_TYPE

{attribute 'external_name' := 'cmp_rts_DFC_MOXEMM_SMU_ALM10_21'}
TYPE DFC_MOXEMM_SMU_ALM10_21 : STRUCT
  DTC : UDINT := 16#10C400;
  DFCid : UINT := 896;
  debounceMethod : USINT := NATIVE;
END_STRUCT;
END_TYPE

{attribute 'external_name' := 'cmp_rts_DFC_MOXEMM_SMU_ALM6_5'}
TYPE DFC_MOXEMM_SMU_ALM6_5 : STRUCT
  DTC : UDINT := 16#109600;
  DFCid : UINT := 957;
  debounceMethod : USINT := NATIVE;
END_STRUCT;
END_TYPE

{attribute 'external_name' := 'cmp_rts_DFC_MOXEMM_SMU_ALM6_7'}
TYPE DFC_MOXEMM_SMU_ALM6_7 : STRUCT
  DTC : UDINT := 16#109700;
  DFCid : UINT := 958;
  debounceMethod : USINT := NATIVE;
END_STRUCT;
END_TYPE

{attribute 'external_name' := 'cmp_rts_DFC_MOXEMM_SMU_ALM6_8'}
TYPE DFC_MOXEMM_SMU_ALM6_8 : STRUCT
  DTC : UDINT := 16#109800;
  DFCid : UINT := 959;
  debounceMethod : USINT := NATIVE;
END_STRUCT;
END_TYPE

{attribute 'external_name' := 'cmp_rts_DFC_COMM_E_NET_START_IND_CHANNEL_3'}
TYPE DFC_COMM_E_NET_START_IND_CHANNEL_3 : STRUCT
  DTC : UDINT := 16#105300;
  DFCid : UINT := 865;
  debounceMethod : USINT := NO_DEBOUNCE;
END_STRUCT;
END_TYPE

{attribute 'external_name' := 'cmp_rts_DFC_COMM_E_NET_START_IND_CHANNEL_2'}
TYPE DFC_COMM_E_NET_START_IND_CHANNEL_2 : STRUCT
  DTC : UDINT := 16#105200;
  DFCid : UINT := 864;
  debounceMethod : USINT := NO_DEBOUNCE;
END_STRUCT;
END_TYPE

{attribute 'external_name' := 'cmp_rts_DFC_COMM_E_NET_START_IND_CHANNEL_5'}
TYPE DFC_COMM_E_NET_START_IND_CHANNEL_5 : STRUCT
  DTC : UDINT := 16#105500;
  DFCid : UINT := 867;
  debounceMethod : USINT := NO_DEBOUNCE;
END_STRUCT;
END_TYPE

{attribute 'external_name' := 'cmp_rts_DFC_COMM_E_NET_START_IND_CHANNEL_4'}
TYPE DFC_COMM_E_NET_START_IND_CHANNEL_4 : STRUCT
  DTC : UDINT := 16#105400;
  DFCid : UINT := 866;
  debounceMethod : USINT := NO_DEBOUNCE;
END_STRUCT;
END_TYPE

{attribute 'external_name' := 'cmp_rts_DFC_MOXEMM_SMU_ALM6_0'}
TYPE DFC_MOXEMM_SMU_ALM6_0 : STRUCT
  DTC : UDINT := 16#109400;
  DFCid : UINT := 945;
  debounceMethod : USINT := NATIVE;
END_STRUCT;
END_TYPE

{attribute 'external_name' := 'cmp_rts_DFC_MOXEMM_SMU_ALM6_2'}
TYPE DFC_MOXEMM_SMU_ALM6_2 : STRUCT
  DTC : UDINT := 16#10D900;
  DFCid : UINT := 952;
  debounceMethod : USINT := NATIVE;
END_STRUCT;
END_TYPE

{attribute 'external_name' := 'cmp_rts_DFC_MOXEMM_SMU_ALM6_4'}
TYPE DFC_MOXEMM_SMU_ALM6_4 : STRUCT
  DTC : UDINT := 16#109500;
  DFCid : UINT := 956;
  debounceMethod : USINT := NATIVE;
END_STRUCT;
END_TYPE

{attribute 'external_name' := 'cmp_rts_DFC_ComCntESP_20'}
TYPE DFC_ComCntESP_20 : STRUCT
  DTC : UDINT := 16#102600;
END_STRUCT;
END_TYPE

{attribute 'external_name' := 'cmp_rts_DFC_ComCntESP_21'}
TYPE DFC_ComCntESP_21 : STRUCT
  DTC : UDINT := 16#102700;
END_STRUCT;
END_TYPE

{attribute 'external_name' := 'cmp_rts_DFC_COMM_E_NET_START_IND_CHANNEL_1'}
TYPE DFC_COMM_E_NET_START_IND_CHANNEL_1 : STRUCT
  DTC : UDINT := 16#105100;
  DFCid : UINT := 863;
  debounceMethod : USINT := NO_DEBOUNCE;
END_STRUCT;
END_TYPE

{attribute 'external_name' := 'cmp_rts_DFC_COMM_E_NET_START_IND_CHANNEL_0'}
TYPE DFC_COMM_E_NET_START_IND_CHANNEL_0 : STRUCT
  DTC : UDINT := 16#105000;
  DFCid : UINT := 862;
  debounceMethod : USINT := NO_DEBOUNCE;
END_STRUCT;
END_TYPE

{attribute 'external_name' := 'cmp_rts_DFC_MOXEMM_SMU_ALM21_0'}
TYPE DFC_MOXEMM_SMU_ALM21_0 : STRUCT
  DTC : UDINT := 16#10CD00;
  DFCid : UINT := 918;
  debounceMethod : USINT := NATIVE;
END_STRUCT;
END_TYPE

{attribute 'external_name' := 'cmp_rts_DFC_MoCSOPICO'}
TYPE DFC_MoCSOPICO : STRUCT
  DTC : UDINT := 16#106000;
  DFCid : UINT := 992;
  debounceMethod : USINT := NATIVE;
END_STRUCT;
END_TYPE

{attribute 'external_name' := 'cmp_rts_DFC_MOXEMM_SMU_ALM21_3'}
TYPE DFC_MOXEMM_SMU_ALM21_3 : STRUCT
  DTC : UDINT := 16#10CE00;
  DFCid : UINT := 920;
  debounceMethod : USINT := NATIVE;
END_STRUCT;
END_TYPE

{attribute 'external_name' := 'cmp_rts_DFC_MoSysCtrlReIni'}
TYPE DFC_MoSysCtrlReIni : STRUCT
  DTC : UDINT := 16#106100;
  DFCid : UINT := 994;
  debounceMethod : USINT := NATIVE;
END_STRUCT;
END_TYPE

{attribute 'external_name' := 'cmp_rts_DFC_RBA_IOEXTLIB_KEEPALIVE_DRV'}
TYPE DFC_RBA_IOEXTLIB_KEEPALIVE_DRV : STRUCT
  DTC : UDINT := 16#094300;
  DFCid : UINT := 871;
  debounceMethod : USINT := NO_DEBOUNCE;
END_STRUCT;
END_TYPE

{attribute 'external_name' := 'cmp_rts_DFC_ComChksESP_20'}
TYPE DFC_ComChksESP_20 : STRUCT
  DTC : UDINT := 16#101D00;
END_STRUCT;
END_TYPE

{attribute 'external_name' := 'cmp_rts_DFC_ComChksESP_21'}
TYPE DFC_ComChksESP_21 : STRUCT
  DTC : UDINT := 16#101E00;
END_STRUCT;
END_TYPE

{attribute 'external_name' := 'cmp_rts_DFC_bds_TimeUpDownDebFault'}
TYPE DFC_bds_TimeUpDownDebFault : STRUCT
  DTC : UDINT := 16#800000;
  DFCid : UINT := 5;
  debounceMethod : USINT := TIME_UP_DOWN;
END_STRUCT;
END_TYPE

{attribute 'external_name' := 'cmp_rts_DFC_bds_EventUpDownDebFault'}
TYPE DFC_bds_EventUpDownDebFault : STRUCT
  DTC : UDINT := 16#800100;
  DFCid : UINT := 517;
  debounceMethod : USINT := EVENT_UP_DOWN;
END_STRUCT;
END_TYPE

{attribute 'external_name' := 'cmp_rts_DFC_bds_EventInRowDebFault'}
TYPE DFC_bds_EventInRowDebFault : STRUCT
  DTC : UDINT := 16#800200;
  DFCid : UINT := 2;
  debounceMethod : USINT := EVENT_IN_ROW;
END_STRUCT;
END_TYPE

{attribute 'external_name' := 'cmp_rts_DFC_bds_TimeInRowDebFault'}
TYPE DFC_bds_TimeInRowDebFault : STRUCT
  DTC : UDINT := 16#800300;
  DFCid : UINT := 1;
  debounceMethod : USINT := TIME_IN_ROW;
END_STRUCT;
END_TYPE

{attribute 'external_name' := 'cmp_rts_DFC_bds_NoDebFault1'}
TYPE DFC_bds_NoDebFault1 : STRUCT
  DTC : UDINT := 16#800400;
  DFCid : UINT := 1007;
  debounceMethod : USINT := NATIVE;
END_STRUCT;
END_TYPE

VAR_GLOBAL  (* GVL_debounceMethod *)
  TIME_IN_ROW : USINT := 0;
  EVENT_IN_ROW : USINT := 1;
  TIME_UP_DOWN : USINT := 2;
  EVENT_UP_DOWN : USINT := 3;
  TIME_UP_DOWN_SMALL : USINT := 4;
  EVENT_UP_DOWN_SMALL : USINT := 5;
  TIME_IN_ROW_SMALL : USINT := 6;
  EVENT_IN_ROW_SMALL : USINT := 7;
  NO_DEBOUNCE : USINT := 8;
  NATIVE : USINT := 8;
END_VAR
